// --- Siemens Structured Format ---
DATA_BLOCK "model__HS32_IW100_"
{ S7_Optimized_Access := 'TRUE' }
VERSION :
NON_RETAIN
   VAR
      W_i : ARRAY[0..31, 0..39] OF REAL;
      W_f : ARRAY[0..31, 0..39] OF REAL;
      W_g : ARRAY[0..31, 0..39] OF REAL;
      W_o : ARRAY[0..31, 0..39] OF REAL;
      R_i : ARRAY[0..31, 0..31] OF REAL;
      R_f : ARRAY[0..31, 0..31] OF REAL;
      R_g : ARRAY[0..31, 0..31] OF REAL;
      R_o : ARRAY[0..31, 0..31] OF REAL;
      B_i : ARRAY[0..31] OF REAL;
      B_f : ARRAY[0..31] OF REAL;
      B_g : ARRAY[0..31] OF REAL;
      B_o : ARRAY[0..31] OF REAL;
      FC_W : ARRAY[0..39, 0..31] OF REAL;
      FC_B : ARRAY[0..39] OF REAL;
   END_VAR
BEGIN

      W_i[0,0] := 0.06179943;
      W_i[0,1] := 0.02775717;
      W_i[0,2] := -0.03196508;
      W_i[0,3] := 0.03677268;
      W_i[0,4] := 0.05541879;
      W_i[0,5] := -0.02846526;
      W_i[0,6] := 0.05010877;
      W_i[0,7] := 0.04675795;
      W_i[0,8] := 0.08269168;
      W_i[0,9] := -0.01895206;
      W_i[0,10] := 0.01859271;
      W_i[0,11] := -0.13412605;
      W_i[0,12] := 0.22322017;
      W_i[0,13] := 0.00698021;
      W_i[0,14] := 0.01548957;
      W_i[0,15] := -0.04365166;
      W_i[0,16] := -0.03781708;
      W_i[0,17] := 0.00911400;
      W_i[0,18] := -0.02057064;
      W_i[0,19] := -0.08685457;
      W_i[0,20] := -0.01680454;
      W_i[0,21] := -0.04614456;
      W_i[0,22] := -0.03545121;
      W_i[0,23] := -0.02339789;
      W_i[0,24] := -1.12611961;
      W_i[0,25] := -0.10453429;
      W_i[0,26] := -0.07026759;
      W_i[0,27] := -0.05480277;
      W_i[0,28] := -0.02404995;
      W_i[0,29] := 0.12750483;
      W_i[0,30] := 0.17675591;
      W_i[0,31] := -0.02635767;
      W_i[0,32] := 0.19571228;
      W_i[0,33] := 0.06735895;
      W_i[0,34] := -0.14900623;
      W_i[0,35] := 0.06775700;
      W_i[0,36] := -0.00490537;
      W_i[0,37] := -0.01378909;
      W_i[0,38] := 0.07458769;
      W_i[0,39] := 0.66414231;
      W_i[1,0] := 0.02071806;
      W_i[1,1] := -0.03353070;
      W_i[1,2] := -0.01928122;
      W_i[1,3] := 0.06214599;
      W_i[1,4] := 0.25778303;
      W_i[1,5] := 0.16688786;
      W_i[1,6] := 0.11954694;
      W_i[1,7] := 0.06900051;
      W_i[1,8] := 0.01723209;
      W_i[1,9] := -0.11005860;
      W_i[1,10] := -0.04237102;
      W_i[1,11] := 0.01513118;
      W_i[1,12] := -0.15226158;
      W_i[1,13] := 0.03596478;
      W_i[1,14] := 0.02140439;
      W_i[1,15] := 0.06197662;
      W_i[1,16] := 0.00865395;
      W_i[1,17] := 0.04867539;
      W_i[1,18] := 0.04397345;
      W_i[1,19] := 0.06557351;
      W_i[1,20] := 0.06942460;
      W_i[1,21] := 0.05065425;
      W_i[1,22] := 0.10510546;
      W_i[1,23] := 0.04281416;
      W_i[1,24] := -0.29392853;
      W_i[1,25] := -0.38343686;
      W_i[1,26] := -0.10036848;
      W_i[1,27] := -0.04264174;
      W_i[1,28] := -0.17839937;
      W_i[1,29] := -0.21495967;
      W_i[1,30] := -0.22097401;
      W_i[1,31] := 0.03829467;
      W_i[1,32] := -0.31760472;
      W_i[1,33] := -0.17684405;
      W_i[1,34] := -0.23336750;
      W_i[1,35] := -0.15993148;
      W_i[1,36] := -0.00517801;
      W_i[1,37] := -0.01187338;
      W_i[1,38] := -0.03392988;
      W_i[1,39] := -0.04533037;
      W_i[2,0] := -0.00829509;
      W_i[2,1] := -0.14865589;
      W_i[2,2] := -0.01495113;
      W_i[2,3] := 0.02128208;
      W_i[2,4] := 0.21340890;
      W_i[2,5] := -0.05039188;
      W_i[2,6] := 0.02410355;
      W_i[2,7] := -0.16800745;
      W_i[2,8] := -0.07282868;
      W_i[2,9] := -0.06157869;
      W_i[2,10] := 0.17263004;
      W_i[2,11] := 0.02063438;
      W_i[2,12] := 0.17519112;
      W_i[2,13] := -0.00622400;
      W_i[2,14] := 0.06819141;
      W_i[2,15] := 0.06226488;
      W_i[2,16] := -0.03465794;
      W_i[2,17] := 0.02215759;
      W_i[2,18] := -0.05341673;
      W_i[2,19] := -0.13253070;
      W_i[2,20] := 0.04460967;
      W_i[2,21] := 0.11263417;
      W_i[2,22] := 0.09742771;
      W_i[2,23] := 0.00662358;
      W_i[2,24] := -0.05392387;
      W_i[2,25] := -0.17852309;
      W_i[2,26] := 0.03923597;
      W_i[2,27] := -0.02955864;
      W_i[2,28] := 0.03645090;
      W_i[2,29] := -0.03638797;
      W_i[2,30] := 0.33836386;
      W_i[2,31] := 0.12495890;
      W_i[2,32] := 0.06078594;
      W_i[2,33] := -0.14091927;
      W_i[2,34] := 0.17067178;
      W_i[2,35] := -0.12043836;
      W_i[2,36] := -0.01742014;
      W_i[2,37] := -0.29951882;
      W_i[2,38] := 0.04487922;
      W_i[2,39] := -0.04771054;
      W_i[3,0] := -0.00100313;
      W_i[3,1] := -0.00449658;
      W_i[3,2] := -0.07554256;
      W_i[3,3] := -0.18185882;
      W_i[3,4] := -0.02607848;
      W_i[3,5] := -0.07896423;
      W_i[3,6] := 0.05784221;
      W_i[3,7] := -0.07038090;
      W_i[3,8] := 0.20566469;
      W_i[3,9] := 0.09180041;
      W_i[3,10] := 0.05098312;
      W_i[3,11] := 0.15374708;
      W_i[3,12] := -0.45315537;
      W_i[3,13] := 0.08420219;
      W_i[3,14] := -0.12126628;
      W_i[3,15] := -0.08021345;
      W_i[3,16] := -0.27470666;
      W_i[3,17] := 0.07300078;
      W_i[3,18] := 0.22311375;
      W_i[3,19] := -0.02914955;
      W_i[3,20] := -0.01066327;
      W_i[3,21] := -0.00681991;
      W_i[3,22] := 0.24156007;
      W_i[3,23] := -0.11151634;
      W_i[3,24] := -0.08966236;
      W_i[3,25] := 0.01983345;
      W_i[3,26] := -0.08444024;
      W_i[3,27] := 0.16410163;
      W_i[3,28] := -0.04299213;
      W_i[3,29] := -0.12410518;
      W_i[3,30] := 0.26584405;
      W_i[3,31] := -0.29169789;
      W_i[3,32] := 0.05328545;
      W_i[3,33] := -0.51094949;
      W_i[3,34] := 0.03447641;
      W_i[3,35] := 0.00506896;
      W_i[3,36] := 0.03782123;
      W_i[3,37] := 0.18697615;
      W_i[3,38] := 0.00981322;
      W_i[3,39] := 0.75137496;
      W_i[4,0] := 0.04553370;
      W_i[4,1] := 0.11792795;
      W_i[4,2] := -0.01621435;
      W_i[4,3] := -0.03620827;
      W_i[4,4] := -0.15278673;
      W_i[4,5] := -0.01032144;
      W_i[4,6] := 0.00459723;
      W_i[4,7] := 0.03891215;
      W_i[4,8] := -0.05662930;
      W_i[4,9] := -0.06458510;
      W_i[4,10] := 0.27832294;
      W_i[4,11] := 0.05678938;
      W_i[4,12] := 0.01970386;
      W_i[4,13] := 0.09437083;
      W_i[4,14] := -0.01984982;
      W_i[4,15] := -0.05285306;
      W_i[4,16] := 0.02962786;
      W_i[4,17] := 0.00963242;
      W_i[4,18] := 0.00985712;
      W_i[4,19] := -0.07215877;
      W_i[4,20] := 0.09223086;
      W_i[4,21] := -0.08452385;
      W_i[4,22] := -0.03868546;
      W_i[4,23] := -0.02803059;
      W_i[4,24] := 0.19232845;
      W_i[4,25] := 0.21442333;
      W_i[4,26] := -0.10829803;
      W_i[4,27] := 0.09679998;
      W_i[4,28] := -0.05681482;
      W_i[4,29] := 0.04554670;
      W_i[4,30] := -0.12465099;
      W_i[4,31] := 0.02753920;
      W_i[4,32] := 0.05632669;
      W_i[4,33] := 0.24204549;
      W_i[4,34] := 0.14613600;
      W_i[4,35] := -0.21246302;
      W_i[4,36] := -0.06815854;
      W_i[4,37] := -0.23073821;
      W_i[4,38] := 0.02998499;
      W_i[4,39] := -0.02546969;
      W_i[5,0] := -0.09215746;
      W_i[5,1] := -0.08727002;
      W_i[5,2] := 0.02556904;
      W_i[5,3] := 0.15369390;
      W_i[5,4] := 0.01142898;
      W_i[5,5] := -0.05077455;
      W_i[5,6] := -0.11507938;
      W_i[5,7] := -0.10518788;
      W_i[5,8] := -0.04785325;
      W_i[5,9] := -0.05123279;
      W_i[5,10] := 0.15905567;
      W_i[5,11] := 0.06097380;
      W_i[5,12] := -0.18418492;
      W_i[5,13] := -0.03047887;
      W_i[5,14] := 0.11933848;
      W_i[5,15] := -0.03554063;
      W_i[5,16] := -0.07242216;
      W_i[5,17] := 0.02859983;
      W_i[5,18] := -0.03490715;
      W_i[5,19] := 0.05818025;
      W_i[5,20] := -0.07515050;
      W_i[5,21] := 0.02579406;
      W_i[5,22] := -0.31216845;
      W_i[5,23] := 0.04713825;
      W_i[5,24] := -0.20269118;
      W_i[5,25] := 0.10239060;
      W_i[5,26] := -0.01558112;
      W_i[5,27] := 0.00159392;
      W_i[5,28] := -0.05441242;
      W_i[5,29] := 0.52095068;
      W_i[5,30] := -0.57061511;
      W_i[5,31] := 0.13902861;
      W_i[5,32] := -0.12816451;
      W_i[5,33] := 0.06774098;
      W_i[5,34] := -0.41744006;
      W_i[5,35] := 0.05064213;
      W_i[5,36] := -0.09991191;
      W_i[5,37] := -0.17586561;
      W_i[5,38] := 0.19242531;
      W_i[5,39] := 0.03359242;
      W_i[6,0] := -0.03353223;
      W_i[6,1] := 0.00677240;
      W_i[6,2] := -0.01104784;
      W_i[6,3] := 0.07707670;
      W_i[6,4] := 0.00404718;
      W_i[6,5] := -0.05442240;
      W_i[6,6] := 0.10070097;
      W_i[6,7] := 0.04808670;
      W_i[6,8] := -0.10168398;
      W_i[6,9] := -0.02940839;
      W_i[6,10] := 0.04046509;
      W_i[6,11] := -0.12609679;
      W_i[6,12] := -0.11311707;
      W_i[6,13] := 0.04389359;
      W_i[6,14] := 0.01754723;
      W_i[6,15] := 0.03694800;
      W_i[6,16] := -0.09526791;
      W_i[6,17] := -0.13010779;
      W_i[6,18] := 0.31546634;
      W_i[6,19] := -0.07569441;
      W_i[6,20] := 0.28956288;
      W_i[6,21] := 0.00949547;
      W_i[6,22] := 0.09859776;
      W_i[6,23] := -0.02917805;
      W_i[6,24] := 0.17138363;
      W_i[6,25] := 0.27182287;
      W_i[6,26] := 0.01862298;
      W_i[6,27] := -0.00405888;
      W_i[6,28] := 0.07469607;
      W_i[6,29] := -0.15340948;
      W_i[6,30] := 0.13516009;
      W_i[6,31] := -0.14186700;
      W_i[6,32] := 0.17514557;
      W_i[6,33] := 0.08133219;
      W_i[6,34] := 0.32842028;
      W_i[6,35] := -0.12072788;
      W_i[6,36] := -0.05676087;
      W_i[6,37] := -0.11963397;
      W_i[6,38] := 0.00256419;
      W_i[6,39] := 0.28269264;
      W_i[7,0] := -0.14775136;
      W_i[7,1] := -0.12126163;
      W_i[7,2] := -0.01920290;
      W_i[7,3] := 0.25063628;
      W_i[7,4] := -0.02222757;
      W_i[7,5] := -0.03862220;
      W_i[7,6] := -0.13837403;
      W_i[7,7] := 0.38717154;
      W_i[7,8] := -0.11613367;
      W_i[7,9] := -0.53373992;
      W_i[7,10] := -0.09174719;
      W_i[7,11] := -0.12254320;
      W_i[7,12] := -0.00825407;
      W_i[7,13] := -0.05826338;
      W_i[7,14] := 0.09619932;
      W_i[7,15] := 0.07305111;
      W_i[7,16] := -0.07672185;
      W_i[7,17] := 0.01172826;
      W_i[7,18] := 0.43864861;
      W_i[7,19] := 0.05868300;
      W_i[7,20] := 0.02254522;
      W_i[7,21] := -0.00708780;
      W_i[7,22] := -0.17880507;
      W_i[7,23] := 0.03120665;
      W_i[7,24] := -0.34886146;
      W_i[7,25] := -0.04237240;
      W_i[7,26] := 0.11693397;
      W_i[7,27] := 0.06307583;
      W_i[7,28] := -0.04923550;
      W_i[7,29] := 0.30479616;
      W_i[7,30] := -0.03511298;
      W_i[7,31] := -0.07993785;
      W_i[7,32] := -0.19723724;
      W_i[7,33] := 0.09875282;
      W_i[7,34] := 0.06003888;
      W_i[7,35] := 0.01167319;
      W_i[7,36] := 0.01233812;
      W_i[7,37] := 0.13565342;
      W_i[7,38] := 0.07438924;
      W_i[7,39] := -0.04580714;
      W_i[8,0] := -0.20123592;
      W_i[8,1] := -0.01675500;
      W_i[8,2] := 0.06737890;
      W_i[8,3] := -0.03567418;
      W_i[8,4] := 0.03670733;
      W_i[8,5] := 0.00518049;
      W_i[8,6] := -0.05625178;
      W_i[8,7] := -0.21017089;
      W_i[8,8] := 0.02617608;
      W_i[8,9] := 0.21776345;
      W_i[8,10] := 0.04046187;
      W_i[8,11] := 0.01215424;
      W_i[8,12] := -0.13758895;
      W_i[8,13] := -0.03766741;
      W_i[8,14] := -0.10688125;
      W_i[8,15] := -0.03897357;
      W_i[8,16] := -0.04154058;
      W_i[8,17] := -0.04646260;
      W_i[8,18] := -0.01917167;
      W_i[8,19] := 0.05721129;
      W_i[8,20] := -0.05588107;
      W_i[8,21] := -0.07682938;
      W_i[8,22] := -0.07860053;
      W_i[8,23] := -0.06132534;
      W_i[8,24] := 0.03326328;
      W_i[8,25] := 0.08150295;
      W_i[8,26] := -0.14111993;
      W_i[8,27] := 0.00011063;
      W_i[8,28] := 0.01932795;
      W_i[8,29] := 0.04262755;
      W_i[8,30] := 0.05650154;
      W_i[8,31] := -0.15539150;
      W_i[8,32] := 0.17859717;
      W_i[8,33] := 0.01948488;
      W_i[8,34] := 0.08800947;
      W_i[8,35] := 0.09776416;
      W_i[8,36] := -0.05269374;
      W_i[8,37] := 0.06550130;
      W_i[8,38] := -0.08607090;
      W_i[8,39] := 0.15070331;
      W_i[9,0] := -0.27159375;
      W_i[9,1] := -0.02797615;
      W_i[9,2] := -0.00100640;
      W_i[9,3] := 0.12800276;
      W_i[9,4] := -0.09242823;
      W_i[9,5] := 0.01892278;
      W_i[9,6] := -0.02738959;
      W_i[9,7] := 0.09567204;
      W_i[9,8] := -0.44594380;
      W_i[9,9] := 0.20733841;
      W_i[9,10] := -0.07766859;
      W_i[9,11] := -0.13440070;
      W_i[9,12] := 0.01596364;
      W_i[9,13] := 0.07334067;
      W_i[9,14] := 0.07882207;
      W_i[9,15] := 0.05607220;
      W_i[9,16] := -0.07642873;
      W_i[9,17] := 0.08819333;
      W_i[9,18] := 0.02835996;
      W_i[9,19] := 0.09605386;
      W_i[9,20] := 0.12935719;
      W_i[9,21] := -0.04795177;
      W_i[9,22] := -0.05849212;
      W_i[9,23] := -0.00860680;
      W_i[9,24] := -0.05882631;
      W_i[9,25] := 0.12313552;
      W_i[9,26] := -0.10078515;
      W_i[9,27] := 0.10558646;
      W_i[9,28] := 0.04912272;
      W_i[9,29] := -0.09551237;
      W_i[9,30] := -0.09409142;
      W_i[9,31] := -0.22199608;
      W_i[9,32] := 0.08531553;
      W_i[9,33] := -0.01295959;
      W_i[9,34] := 0.28744900;
      W_i[9,35] := -0.14239824;
      W_i[9,36] := -0.16849788;
      W_i[9,37] := -0.06152735;
      W_i[9,38] := 0.01881091;
      W_i[9,39] := -0.08872003;
      W_i[10,0] := 0.04977950;
      W_i[10,1] := 0.01497823;
      W_i[10,2] := -0.00536506;
      W_i[10,3] := 0.02952771;
      W_i[10,4] := -0.03139960;
      W_i[10,5] := -0.00463935;
      W_i[10,6] := -0.10389712;
      W_i[10,7] := -0.10033682;
      W_i[10,8] := 0.11073951;
      W_i[10,9] := -0.08885644;
      W_i[10,10] := 0.01201617;
      W_i[10,11] := -0.63600385;
      W_i[10,12] := 0.57826489;
      W_i[10,13] := -0.00285191;
      W_i[10,14] := -0.13222906;
      W_i[10,15] := 0.01793578;
      W_i[10,16] := -0.03972865;
      W_i[10,17] := 0.16141385;
      W_i[10,18] := 0.48685026;
      W_i[10,19] := -0.04842542;
      W_i[10,20] := 0.03557721;
      W_i[10,21] := -0.02083956;
      W_i[10,22] := 0.07665567;
      W_i[10,23] := 0.13016869;
      W_i[10,24] := -0.08724608;
      W_i[10,25] := -0.20036544;
      W_i[10,26] := -0.12496603;
      W_i[10,27] := -0.05189490;
      W_i[10,28] := 0.10159702;
      W_i[10,29] := -0.05331298;
      W_i[10,30] := 0.03033962;
      W_i[10,31] := 0.07102174;
      W_i[10,32] := 0.02948349;
      W_i[10,33] := 0.01139331;
      W_i[10,34] := -0.43736589;
      W_i[10,35] := 0.28173751;
      W_i[10,36] := 0.01866223;
      W_i[10,37] := 0.25957814;
      W_i[10,38] := 0.14778605;
      W_i[10,39] := 0.93045533;
      W_i[11,0] := -0.10133153;
      W_i[11,1] := -0.05051550;
      W_i[11,2] := -0.03669089;
      W_i[11,3] := 0.14228435;
      W_i[11,4] := 0.08680110;
      W_i[11,5] := 0.02299375;
      W_i[11,6] := -0.11019665;
      W_i[11,7] := 0.03878751;
      W_i[11,8] := 0.05327412;
      W_i[11,9] := -0.29215959;
      W_i[11,10] := -0.06103910;
      W_i[11,11] := -0.04436091;
      W_i[11,12] := 0.10810567;
      W_i[11,13] := -0.12327234;
      W_i[11,14] := -0.03792057;
      W_i[11,15] := -0.01659554;
      W_i[11,16] := 0.01878507;
      W_i[11,17] := -0.00647482;
      W_i[11,18] := -0.04410561;
      W_i[11,19] := 0.07929806;
      W_i[11,20] := 0.01020784;
      W_i[11,21] := 0.08437648;
      W_i[11,22] := 0.10375391;
      W_i[11,23] := 0.20762387;
      W_i[11,24] := -0.57340568;
      W_i[11,25] := -0.59531760;
      W_i[11,26] := -0.17425776;
      W_i[11,27] := -0.11098373;
      W_i[11,28] := 0.01483229;
      W_i[11,29] := 0.08123992;
      W_i[11,30] := 0.16729805;
      W_i[11,31] := -0.17426890;
      W_i[11,32] := 0.17722335;
      W_i[11,33] := -0.07652548;
      W_i[11,34] := 0.18267493;
      W_i[11,35] := 0.19876397;
      W_i[11,36] := 0.04698262;
      W_i[11,37] := 0.02095936;
      W_i[11,38] := -0.10085329;
      W_i[11,39] := 1.06740248;
      W_i[12,0] := -0.12894745;
      W_i[12,1] := -0.01604900;
      W_i[12,2] := -0.05750192;
      W_i[12,3] := 0.08071270;
      W_i[12,4] := -0.10707285;
      W_i[12,5] := -0.09226165;
      W_i[12,6] := 0.01451022;
      W_i[12,7] := 0.16588750;
      W_i[12,8] := -0.20528767;
      W_i[12,9] := 0.16444704;
      W_i[12,10] := 0.09167138;
      W_i[12,11] := -0.05738107;
      W_i[12,12] := -0.03085519;
      W_i[12,13] := 0.02227092;
      W_i[12,14] := 0.00619229;
      W_i[12,15] := 0.07799102;
      W_i[12,16] := 0.02899228;
      W_i[12,17] := 0.01908563;
      W_i[12,18] := 0.55716008;
      W_i[12,19] := 0.09226023;
      W_i[12,20] := -0.01587960;
      W_i[12,21] := -0.13448635;
      W_i[12,22] := -0.14700012;
      W_i[12,23] := -0.06094320;
      W_i[12,24] := 0.27282214;
      W_i[12,25] := 0.21529709;
      W_i[12,26] := -0.12392846;
      W_i[12,27] := 0.05751082;
      W_i[12,28] := 0.12284551;
      W_i[12,29] := -0.00490399;
      W_i[12,30] := -0.17141145;
      W_i[12,31] := -0.08434223;
      W_i[12,32] := 0.05438624;
      W_i[12,33] := -0.10759345;
      W_i[12,34] := -0.07436828;
      W_i[12,35] := -0.12592168;
      W_i[12,36] := 0.02604092;
      W_i[12,37] := -0.15142396;
      W_i[12,38] := -0.03170886;
      W_i[12,39] := 0.16621175;
      W_i[13,0] := -0.00913993;
      W_i[13,1] := -0.04174744;
      W_i[13,2] := -0.03129856;
      W_i[13,3] := -0.04003599;
      W_i[13,4] := 0.04255468;
      W_i[13,5] := 0.00480728;
      W_i[13,6] := -0.07061405;
      W_i[13,7] := -0.03280373;
      W_i[13,8] := 0.02827574;
      W_i[13,9] := 0.02418965;
      W_i[13,10] := 0.07189363;
      W_i[13,11] := 0.12613529;
      W_i[13,12] := 0.03361855;
      W_i[13,13] := 0.03988501;
      W_i[13,14] := -0.02885863;
      W_i[13,15] := -0.00470651;
      W_i[13,16] := -0.03359226;
      W_i[13,17] := -0.00056631;
      W_i[13,18] := -0.07915758;
      W_i[13,19] := 0.01315921;
      W_i[13,20] := 0.10718971;
      W_i[13,21] := 0.13062805;
      W_i[13,22] := 0.16784896;
      W_i[13,23] := -0.07162543;
      W_i[13,24] := 0.03916876;
      W_i[13,25] := -0.11025614;
      W_i[13,26] := -0.04175865;
      W_i[13,27] := -0.27723673;
      W_i[13,28] := 0.18863167;
      W_i[13,29] := 0.18414941;
      W_i[13,30] := 0.21448347;
      W_i[13,31] := 0.27937597;
      W_i[13,32] := -0.15358151;
      W_i[13,33] := 0.04613268;
      W_i[13,34] := -0.28416333;
      W_i[13,35] := -0.24947314;
      W_i[13,36] := -0.06312902;
      W_i[13,37] := -0.19301520;
      W_i[13,38] := 0.07415584;
      W_i[13,39] := 0.07214847;
      W_i[14,0] := -0.06886686;
      W_i[14,1] := 0.09983595;
      W_i[14,2] := 0.00539746;
      W_i[14,3] := 0.03236075;
      W_i[14,4] := 0.30145952;
      W_i[14,5] := 0.10646193;
      W_i[14,6] := -0.00687617;
      W_i[14,7] := -0.02083724;
      W_i[14,8] := 0.09362940;
      W_i[14,9] := 0.24021219;
      W_i[14,10] := -0.51702040;
      W_i[14,11] := 0.00785133;
      W_i[14,12] := -0.06570137;
      W_i[14,13] := 0.00066462;
      W_i[14,14] := 0.04833549;
      W_i[14,15] := 0.01324825;
      W_i[14,16] := 0.00547472;
      W_i[14,17] := 0.03968929;
      W_i[14,18] := -0.05878792;
      W_i[14,19] := -0.12701105;
      W_i[14,20] := 0.64508420;
      W_i[14,21] := -0.02393116;
      W_i[14,22] := 0.01463204;
      W_i[14,23] := 0.09599538;
      W_i[14,24] := -0.01352467;
      W_i[14,25] := -0.09434310;
      W_i[14,26] := 0.09360847;
      W_i[14,27] := 0.19543391;
      W_i[14,28] := -0.08615168;
      W_i[14,29] := 0.51883084;
      W_i[14,30] := 0.05632273;
      W_i[14,31] := 0.31189725;
      W_i[14,32] := -0.08525938;
      W_i[14,33] := 0.18389013;
      W_i[14,34] := 0.22316632;
      W_i[14,35] := -0.11821964;
      W_i[14,36] := 0.02146083;
      W_i[14,37] := -0.16101155;
      W_i[14,38] := 0.00918483;
      W_i[14,39] := -0.08109198;
      W_i[15,0] := 0.08172593;
      W_i[15,1] := -0.15062873;
      W_i[15,2] := 0.00789237;
      W_i[15,3] := -0.12266801;
      W_i[15,4] := -0.01449642;
      W_i[15,5] := -0.08026960;
      W_i[15,6] := 0.00158959;
      W_i[15,7] := -0.17118339;
      W_i[15,8] := 0.06299323;
      W_i[15,9] := 0.08208384;
      W_i[15,10] := 0.04913726;
      W_i[15,11] := -0.04209859;
      W_i[15,12] := 0.14104722;
      W_i[15,13] := 0.08269731;
      W_i[15,14] := -0.00785436;
      W_i[15,15] := 0.01761792;
      W_i[15,16] := 0.06018753;
      W_i[15,17] := 0.01103730;
      W_i[15,18] := 0.60089856;
      W_i[15,19] := -0.02956709;
      W_i[15,20] := -0.06978408;
      W_i[15,21] := -0.10184263;
      W_i[15,22] := -0.08161820;
      W_i[15,23] := -0.09385420;
      W_i[15,24] := -0.25269318;
      W_i[15,25] := -0.36792046;
      W_i[15,26] := -0.02104633;
      W_i[15,27] := 0.08724175;
      W_i[15,28] := -0.02899375;
      W_i[15,29] := 0.06102180;
      W_i[15,30] := -0.07059706;
      W_i[15,31] := 0.02143796;
      W_i[15,32] := -0.10914523;
      W_i[15,33] := -0.00082962;
      W_i[15,34] := -0.13892201;
      W_i[15,35] := 0.03998528;
      W_i[15,36] := -0.00446972;
      W_i[15,37] := 0.06410963;
      W_i[15,38] := -0.09802709;
      W_i[15,39] := 0.13650982;
      W_i[16,0] := 0.00692594;
      W_i[16,1] := -0.06901163;
      W_i[16,2] := -0.06960113;
      W_i[16,3] := 0.01490095;
      W_i[16,4] := 0.11437556;
      W_i[16,5] := -0.10528261;
      W_i[16,6] := 0.06423379;
      W_i[16,7] := -0.09478712;
      W_i[16,8] := -0.00620357;
      W_i[16,9] := 0.04550839;
      W_i[16,10] := 0.06371807;
      W_i[16,11] := -0.22288436;
      W_i[16,12] := 0.11317084;
      W_i[16,13] := -0.00150014;
      W_i[16,14] := 0.03941125;
      W_i[16,15] := 0.23517418;
      W_i[16,16] := 0.06774591;
      W_i[16,17] := -0.06179966;
      W_i[16,18] := -0.02661809;
      W_i[16,19] := -0.46718821;
      W_i[16,20] := 0.00290592;
      W_i[16,21] := 0.08730330;
      W_i[16,22] := -0.17280819;
      W_i[16,23] := 0.04183443;
      W_i[16,24] := -0.15965074;
      W_i[16,25] := -0.21877262;
      W_i[16,26] := 0.03479860;
      W_i[16,27] := -0.03698987;
      W_i[16,28] := -0.04753701;
      W_i[16,29] := 0.12801097;
      W_i[16,30] := 0.04739811;
      W_i[16,31] := -0.00796509;
      W_i[16,32] := -0.10788697;
      W_i[16,33] := -0.08236082;
      W_i[16,34] := -0.41695821;
      W_i[16,35] := 0.02638846;
      W_i[16,36] := -0.05947839;
      W_i[16,37] := -0.08056837;
      W_i[16,38] := 0.04219051;
      W_i[16,39] := -0.06786148;
      W_i[17,0] := 0.19944434;
      W_i[17,1] := 0.11471956;
      W_i[17,2] := 0.00180160;
      W_i[17,3] := 0.11797725;
      W_i[17,4] := -0.12125240;
      W_i[17,5] := 0.27995679;
      W_i[17,6] := -0.34394604;
      W_i[17,7] := 0.02910547;
      W_i[17,8] := -0.19582599;
      W_i[17,9] := -0.11236304;
      W_i[17,10] := -0.31493005;
      W_i[17,11] := -0.24195738;
      W_i[17,12] := -0.07686605;
      W_i[17,13] := 0.14992486;
      W_i[17,14] := -0.19373207;
      W_i[17,15] := -0.25997469;
      W_i[17,16] := 0.04234881;
      W_i[17,17] := -0.07211331;
      W_i[17,18] := 0.13888460;
      W_i[17,19] := -0.12404422;
      W_i[17,20] := -0.08650170;
      W_i[17,21] := 0.22232069;
      W_i[17,22] := 0.02460083;
      W_i[17,23] := -0.23321719;
      W_i[17,24] := 0.27493891;
      W_i[17,25] := 0.29532185;
      W_i[17,26] := -0.09839682;
      W_i[17,27] := -0.27084854;
      W_i[17,28] := 0.16536197;
      W_i[17,29] := 0.96769738;
      W_i[17,30] := 0.08850956;
      W_i[17,31] := 0.44717026;
      W_i[17,32] := 0.05195052;
      W_i[17,33] := -0.25492772;
      W_i[17,34] := 0.08993755;
      W_i[17,35] := 0.11916504;
      W_i[17,36] := 0.51604098;
      W_i[17,37] := -0.19514880;
      W_i[17,38] := 0.03904369;
      W_i[17,39] := -1.25412786;
      W_i[18,0] := 0.26778793;
      W_i[18,1] := -0.01803258;
      W_i[18,2] := -0.35264796;
      W_i[18,3] := -0.03628552;
      W_i[18,4] := -0.09051698;
      W_i[18,5] := -0.07353226;
      W_i[18,6] := -0.03659349;
      W_i[18,7] := 0.01280040;
      W_i[18,8] := -0.03461934;
      W_i[18,9] := 0.05958343;
      W_i[18,10] := 0.05166731;
      W_i[18,11] := -0.09699293;
      W_i[18,12] := -0.12538935;
      W_i[18,13] := -0.00645365;
      W_i[18,14] := 0.02199500;
      W_i[18,15] := -0.03021014;
      W_i[18,16] := 0.18712366;
      W_i[18,17] := -0.01909142;
      W_i[18,18] := 0.02058483;
      W_i[18,19] := 0.08988243;
      W_i[18,20] := 0.07572187;
      W_i[18,21] := 0.08197203;
      W_i[18,22] := -0.07564746;
      W_i[18,23] := 0.03924798;
      W_i[18,24] := -0.40492132;
      W_i[18,25] := -0.37123427;
      W_i[18,26] := 0.04573231;
      W_i[18,27] := -0.01739427;
      W_i[18,28] := -0.00431714;
      W_i[18,29] := 0.16991295;
      W_i[18,30] := -0.03938163;
      W_i[18,31] := -0.01546910;
      W_i[18,32] := -0.25745204;
      W_i[18,33] := 0.13622859;
      W_i[18,34] := -0.16286966;
      W_i[18,35] := -0.25323087;
      W_i[18,36] := 0.02914849;
      W_i[18,37] := 0.00573681;
      W_i[18,38] := -0.05729824;
      W_i[18,39] := 0.23888165;
      W_i[19,0] := -0.05738360;
      W_i[19,1] := 0.05517812;
      W_i[19,2] := -0.01163843;
      W_i[19,3] := -0.07037261;
      W_i[19,4] := -0.07145417;
      W_i[19,5] := 0.08916121;
      W_i[19,6] := -0.05329772;
      W_i[19,7] := -0.17612284;
      W_i[19,8] := -0.03184425;
      W_i[19,9] := 0.03378281;
      W_i[19,10] := 0.06813814;
      W_i[19,11] := 0.08680203;
      W_i[19,12] := -0.17591415;
      W_i[19,13] := -0.04395442;
      W_i[19,14] := 0.10378881;
      W_i[19,15] := 0.11948365;
      W_i[19,16] := -0.11327706;
      W_i[19,17] := 0.03809229;
      W_i[19,18] := 0.04363121;
      W_i[19,19] := -0.08202547;
      W_i[19,20] := 0.04668652;
      W_i[19,21] := -0.06396332;
      W_i[19,22] := -0.11801164;
      W_i[19,23] := 0.00545785;
      W_i[19,24] := 0.19188444;
      W_i[19,25] := 0.15162137;
      W_i[19,26] := -0.08233768;
      W_i[19,27] := 0.10989103;
      W_i[19,28] := 0.06658027;
      W_i[19,29] := -0.12314930;
      W_i[19,30] := -0.29401505;
      W_i[19,31] := -0.02752479;
      W_i[19,32] := -0.06132220;
      W_i[19,33] := -0.22982699;
      W_i[19,34] := -0.23728208;
      W_i[19,35] := -0.25140384;
      W_i[19,36] := -0.05633686;
      W_i[19,37] := -0.18172039;
      W_i[19,38] := 0.11977114;
      W_i[19,39] := -0.16488980;
      W_i[20,0] := -0.01835487;
      W_i[20,1] := -0.04570545;
      W_i[20,2] := 0.04467667;
      W_i[20,3] := -0.07336899;
      W_i[20,4] := 0.02571872;
      W_i[20,5] := -0.01889678;
      W_i[20,6] := -0.02779749;
      W_i[20,7] := 0.08607043;
      W_i[20,8] := 0.01099925;
      W_i[20,9] := -0.00992060;
      W_i[20,10] := -0.01524233;
      W_i[20,11] := 0.21199150;
      W_i[20,12] := 0.01592732;
      W_i[20,13] := -0.01826751;
      W_i[20,14] := -0.10014486;
      W_i[20,15] := 0.00661277;
      W_i[20,16] := 0.01667893;
      W_i[20,17] := 0.02136482;
      W_i[20,18] := 0.03966679;
      W_i[20,19] := -0.07920662;
      W_i[20,20] := 0.06787179;
      W_i[20,21] := 0.42317262;
      W_i[20,22] := -0.33591220;
      W_i[20,23] := -0.00585524;
      W_i[20,24] := 0.09470745;
      W_i[20,25] := 0.15506293;
      W_i[20,26] := -0.30801183;
      W_i[20,27] := -0.33458385;
      W_i[20,28] := -0.08752628;
      W_i[20,29] := 0.35584134;
      W_i[20,30] := -0.20388263;
      W_i[20,31] := -0.01898901;
      W_i[20,32] := -0.41883579;
      W_i[20,33] := -0.54509979;
      W_i[20,34] := -0.31911835;
      W_i[20,35] := 0.02712717;
      W_i[20,36] := -0.01844929;
      W_i[20,37] := 0.01240083;
      W_i[20,38] := -0.24291822;
      W_i[20,39] := -0.17812274;
      W_i[21,0] := 0.12280829;
      W_i[21,1] := -0.07471990;
      W_i[21,2] := -0.05163937;
      W_i[21,3] := -0.22502938;
      W_i[21,4] := 0.00184776;
      W_i[21,5] := -0.01510628;
      W_i[21,6] := 0.13238980;
      W_i[21,7] := -0.09605303;
      W_i[21,8] := 0.05345604;
      W_i[21,9] := 0.25691971;
      W_i[21,10] := 0.00038861;
      W_i[21,11] := -0.01645699;
      W_i[21,12] := -0.07529693;
      W_i[21,13] := -0.01089604;
      W_i[21,14] := 0.07050634;
      W_i[21,15] := -0.01411841;
      W_i[21,16] := -0.09095489;
      W_i[21,17] := -0.02065623;
      W_i[21,18] := 0.05196851;
      W_i[21,19] := 0.80753618;
      W_i[21,20] := -0.02273143;
      W_i[21,21] := 0.03218904;
      W_i[21,22] := 0.16152497;
      W_i[21,23] := -0.01746419;
      W_i[21,24] := 0.70909500;
      W_i[21,25] := 0.95648199;
      W_i[21,26] := 0.13566963;
      W_i[21,27] := 0.11187585;
      W_i[21,28] := 0.08011223;
      W_i[21,29] := -0.13311587;
      W_i[21,30] := 0.02521890;
      W_i[21,31] := 0.09288229;
      W_i[21,32] := 0.16024679;
      W_i[21,33] := 0.04743494;
      W_i[21,34] := -0.09396220;
      W_i[21,35] := 0.12562209;
      W_i[21,36] := 0.04016363;
      W_i[21,37] := 0.29017061;
      W_i[21,38] := 0.02795759;
      W_i[21,39] := 0.36647096;
      W_i[22,0] := 0.06585112;
      W_i[22,1] := -0.07038485;
      W_i[22,2] := 0.03823679;
      W_i[22,3] := 0.13506269;
      W_i[22,4] := 0.06941289;
      W_i[22,5] := -0.08188840;
      W_i[22,6] := -0.00802410;
      W_i[22,7] := 0.00843967;
      W_i[22,8] := 0.03293480;
      W_i[22,9] := 0.00418619;
      W_i[22,10] := -0.18440005;
      W_i[22,11] := -0.07325464;
      W_i[22,12] := -0.14550987;
      W_i[22,13] := -0.08753653;
      W_i[22,14] := 0.04707590;
      W_i[22,15] := 0.02154654;
      W_i[22,16] := -0.05312854;
      W_i[22,17] := -0.00624513;
      W_i[22,18] := -0.05160676;
      W_i[22,19] := 0.08727906;
      W_i[22,20] := 0.02189743;
      W_i[22,21] := 0.08372616;
      W_i[22,22] := 0.26144525;
      W_i[22,23] := 0.16893846;
      W_i[22,24] := -0.15793604;
      W_i[22,25] := -0.13311699;
      W_i[22,26] := -0.11365860;
      W_i[22,27] := 0.00836681;
      W_i[22,28] := -0.09337366;
      W_i[22,29] := -0.01833472;
      W_i[22,30] := -0.04223403;
      W_i[22,31] := -0.05326389;
      W_i[22,32] := 0.19289488;
      W_i[22,33] := 0.05630151;
      W_i[22,34] := 0.27636716;
      W_i[22,35] := -0.09883546;
      W_i[22,36] := 0.07930394;
      W_i[22,37] := -0.02333659;
      W_i[22,38] := 0.02749063;
      W_i[22,39] := -0.01253646;
      W_i[23,0] := 0.01285714;
      W_i[23,1] := -0.01090977;
      W_i[23,2] := -0.12196957;
      W_i[23,3] := 0.08748322;
      W_i[23,4] := -0.04398613;
      W_i[23,5] := -0.13556443;
      W_i[23,6] := 0.02350867;
      W_i[23,7] := -0.11876588;
      W_i[23,8] := 0.10013366;
      W_i[23,9] := 0.02939740;
      W_i[23,10] := -0.09517333;
      W_i[23,11] := 0.11568693;
      W_i[23,12] := -0.36971363;
      W_i[23,13] := -0.06232831;
      W_i[23,14] := 0.02247390;
      W_i[23,15] := 0.01112311;
      W_i[23,16] := -0.05705897;
      W_i[23,17] := 0.06032606;
      W_i[23,18] := 0.32368115;
      W_i[23,19] := -0.10644881;
      W_i[23,20] := -0.04895338;
      W_i[23,21] := 0.09499650;
      W_i[23,22] := -0.10231195;
      W_i[23,23] := -0.01488803;
      W_i[23,24] := -0.22148487;
      W_i[23,25] := -0.02040800;
      W_i[23,26] := 0.18095909;
      W_i[23,27] := -0.01085224;
      W_i[23,28] := 0.08920502;
      W_i[23,29] := 0.30755806;
      W_i[23,30] := -0.21824111;
      W_i[23,31] := -0.06937134;
      W_i[23,32] := 0.14039119;
      W_i[23,33] := 0.22622369;
      W_i[23,34] := -0.10339716;
      W_i[23,35] := 0.05056783;
      W_i[23,36] := -0.01605630;
      W_i[23,37] := 0.21682332;
      W_i[23,38] := 0.91564023;
      W_i[23,39] := 0.60147935;
      W_i[24,0] := -0.06349316;
      W_i[24,1] := -0.06430539;
      W_i[24,2] := 0.04938103;
      W_i[24,3] := 0.02899365;
      W_i[24,4] := 0.02045459;
      W_i[24,5] := -0.03727232;
      W_i[24,6] := 0.01954682;
      W_i[24,7] := -0.10346385;
      W_i[24,8] := 0.00335618;
      W_i[24,9] := -0.11790799;
      W_i[24,10] := 0.04728369;
      W_i[24,11] := 0.09648414;
      W_i[24,12] := -0.04300074;
      W_i[24,13] := 0.02185826;
      W_i[24,14] := 0.01268934;
      W_i[24,15] := -0.03640975;
      W_i[24,16] := -0.00692598;
      W_i[24,17] := -0.01243239;
      W_i[24,18] := 0.02085917;
      W_i[24,19] := 0.02911621;
      W_i[24,20] := 0.11124941;
      W_i[24,21] := 0.14329974;
      W_i[24,22] := 0.07946618;
      W_i[24,23] := 0.01397222;
      W_i[24,24] := -0.33342758;
      W_i[24,25] := -0.18193676;
      W_i[24,26] := -0.12712136;
      W_i[24,27] := -0.03829253;
      W_i[24,28] := 0.01048399;
      W_i[24,29] := -0.12682118;
      W_i[24,30] := 0.06314925;
      W_i[24,31] := 0.08736062;
      W_i[24,32] := -0.07333044;
      W_i[24,33] := -0.18093891;
      W_i[24,34] := 0.08127785;
      W_i[24,35] := -0.14450674;
      W_i[24,36] := -0.05644464;
      W_i[24,37] := -0.06005542;
      W_i[24,38] := 0.01570564;
      W_i[24,39] := 0.04107951;
      W_i[25,0] := -0.00392134;
      W_i[25,1] := -0.02218844;
      W_i[25,2] := 0.01908197;
      W_i[25,3] := 0.00515596;
      W_i[25,4] := -0.06599259;
      W_i[25,5] := -0.09139763;
      W_i[25,6] := 0.06393541;
      W_i[25,7] := -0.03314249;
      W_i[25,8] := -0.00094995;
      W_i[25,9] := -0.09238666;
      W_i[25,10] := 0.12895916;
      W_i[25,11] := -0.03478534;
      W_i[25,12] := 0.08731889;
      W_i[25,13] := 0.00909062;
      W_i[25,14] := 0.03396220;
      W_i[25,15] := 0.00441095;
      W_i[25,16] := -0.08805312;
      W_i[25,17] := 0.06228795;
      W_i[25,18] := -0.04030024;
      W_i[25,19] := -0.05294413;
      W_i[25,20] := -0.03475821;
      W_i[25,21] := -0.09267792;
      W_i[25,22] := -0.11669731;
      W_i[25,23] := -0.03766777;
      W_i[25,24] := -0.03449144;
      W_i[25,25] := -0.15750119;
      W_i[25,26] := 0.02700294;
      W_i[25,27] := 0.10468993;
      W_i[25,28] := 0.03980485;
      W_i[25,29] := 0.01171093;
      W_i[25,30] := 0.08682661;
      W_i[25,31] := -0.00671425;
      W_i[25,32] := 0.00725360;
      W_i[25,33] := -0.11579906;
      W_i[25,34] := -0.55428278;
      W_i[25,35] := 0.18704750;
      W_i[25,36] := -0.03766178;
      W_i[25,37] := -0.09676717;
      W_i[25,38] := 0.10681428;
      W_i[25,39] := -0.04854197;
      W_i[26,0] := 0.03223363;
      W_i[26,1] := -0.11389477;
      W_i[26,2] := 0.01710660;
      W_i[26,3] := -0.06687164;
      W_i[26,4] := 0.01613229;
      W_i[26,5] := -0.03883494;
      W_i[26,6] := -0.10788758;
      W_i[26,7] := 0.04997331;
      W_i[26,8] := 0.00840330;
      W_i[26,9] := -0.06306913;
      W_i[26,10] := 0.06178190;
      W_i[26,11] := -0.12198523;
      W_i[26,12] := -0.04752781;
      W_i[26,13] := -0.03431008;
      W_i[26,14] := 0.00714531;
      W_i[26,15] := 0.05213116;
      W_i[26,16] := 0.01167048;
      W_i[26,17] := -0.00677893;
      W_i[26,18] := -0.24137808;
      W_i[26,19] := -0.07195701;
      W_i[26,20] := -0.10280736;
      W_i[26,21] := -0.00431173;
      W_i[26,22] := -0.40525341;
      W_i[26,23] := 0.00794029;
      W_i[26,24] := -0.36122626;
      W_i[26,25] := 0.04784513;
      W_i[26,26] := -0.29187959;
      W_i[26,27] := -0.14297174;
      W_i[26,28] := 0.02196433;
      W_i[26,29] := 0.49258694;
      W_i[26,30] := -0.35673437;
      W_i[26,31] := -0.14768223;
      W_i[26,32] := -0.14340006;
      W_i[26,33] := -0.10875791;
      W_i[26,34] := -0.22464323;
      W_i[26,35] := -0.14221328;
      W_i[26,36] := -0.07692026;
      W_i[26,37] := -0.33565632;
      W_i[26,38] := -0.03680801;
      W_i[26,39] := -0.08500476;
      W_i[27,0] := -0.03908358;
      W_i[27,1] := 0.06247386;
      W_i[27,2] := 0.07315844;
      W_i[27,3] := -0.12355068;
      W_i[27,4] := 0.05118919;
      W_i[27,5] := -0.01427916;
      W_i[27,6] := 0.12830800;
      W_i[27,7] := 0.12413668;
      W_i[27,8] := -0.04524078;
      W_i[27,9] := 0.12099374;
      W_i[27,10] := 0.00551115;
      W_i[27,11] := 0.29388657;
      W_i[27,12] := -0.18307312;
      W_i[27,13] := 0.04645123;
      W_i[27,14] := 0.01536438;
      W_i[27,15] := -0.15575469;
      W_i[27,16] := -0.06600323;
      W_i[27,17] := 0.00907420;
      W_i[27,18] := 0.76988453;
      W_i[27,19] := 0.03355170;
      W_i[27,20] := -0.00380640;
      W_i[27,21] := 0.02491378;
      W_i[27,22] := 0.00787842;
      W_i[27,23] := -0.03097626;
      W_i[27,24] := 0.01564326;
      W_i[27,25] := 0.19453372;
      W_i[27,26] := 0.06244323;
      W_i[27,27] := 0.05636120;
      W_i[27,28] := -0.16548483;
      W_i[27,29] := -0.05327202;
      W_i[27,30] := 0.07400166;
      W_i[27,31] := -0.14070928;
      W_i[27,32] := -0.00810295;
      W_i[27,33] := 0.09415199;
      W_i[27,34] := -0.15936106;
      W_i[27,35] := 0.11152661;
      W_i[27,36] := 0.03231200;
      W_i[27,37] := 0.04753703;
      W_i[27,38] := 0.23126490;
      W_i[27,39] := 0.00431150;
      W_i[28,0] := 0.03881709;
      W_i[28,1] := -0.04091561;
      W_i[28,2] := 0.01611770;
      W_i[28,3] := 0.00697450;
      W_i[28,4] := 0.18305339;
      W_i[28,5] := -0.15279785;
      W_i[28,6] := 0.04542335;
      W_i[28,7] := 0.19088306;
      W_i[28,8] := -0.09130806;
      W_i[28,9] := -0.06414899;
      W_i[28,10] := -0.17731205;
      W_i[28,11] := 0.30202127;
      W_i[28,12] := -0.05439992;
      W_i[28,13] := -0.01150446;
      W_i[28,14] := 0.00131535;
      W_i[28,15] := -0.09205615;
      W_i[28,16] := 0.00188813;
      W_i[28,17] := 0.02027261;
      W_i[28,18] := -0.10595226;
      W_i[28,19] := 0.04467888;
      W_i[28,20] := 0.06951932;
      W_i[28,21] := -0.00705112;
      W_i[28,22] := 0.26304314;
      W_i[28,23] := -0.06421968;
      W_i[28,24] := -0.06970753;
      W_i[28,25] := -0.04688016;
      W_i[28,26] := -0.12970042;
      W_i[28,27] := -0.15225610;
      W_i[28,28] := -0.09705786;
      W_i[28,29] := 0.48931244;
      W_i[28,30] := 0.07042009;
      W_i[28,31] := 0.21406028;
      W_i[28,32] := 0.07373387;
      W_i[28,33] := 0.03300231;
      W_i[28,34] := 0.03395164;
      W_i[28,35] := 0.00114277;
      W_i[28,36] := 0.11038067;
      W_i[28,37] := 0.08363102;
      W_i[28,38] := 0.06231136;
      W_i[28,39] := 0.02984152;
      W_i[29,0] := 0.34138203;
      W_i[29,1] := 0.16524114;
      W_i[29,2] := -0.15652245;
      W_i[29,3] := 0.16650911;
      W_i[29,4] := 0.18447480;
      W_i[29,5] := 0.09144969;
      W_i[29,6] := 0.01847808;
      W_i[29,7] := -0.09755348;
      W_i[29,8] := 0.06849403;
      W_i[29,9] := -0.12883465;
      W_i[29,10] := -0.08249056;
      W_i[29,11] := -0.14052261;
      W_i[29,12] := 0.00471857;
      W_i[29,13] := 0.11108005;
      W_i[29,14] := 0.00168034;
      W_i[29,15] := 0.01264171;
      W_i[29,16] := 0.03052950;
      W_i[29,17] := -0.01635699;
      W_i[29,18] := 0.68267095;
      W_i[29,19] := 0.05182270;
      W_i[29,20] := 0.04084420;
      W_i[29,21] := -0.13725121;
      W_i[29,22] := -0.06725579;
      W_i[29,23] := 0.06445967;
      W_i[29,24] := -0.25235596;
      W_i[29,25] := -0.34174517;
      W_i[29,26] := -0.12284433;
      W_i[29,27] := 0.01959689;
      W_i[29,28] := -0.15510176;
      W_i[29,29] := -0.05445927;
      W_i[29,30] := -0.00391692;
      W_i[29,31] := 0.09164531;
      W_i[29,32] := -0.03895570;
      W_i[29,33] := 0.01729037;
      W_i[29,34] := -0.47271654;
      W_i[29,35] := -0.19013441;
      W_i[29,36] := 0.02730786;
      W_i[29,37] := -0.10548180;
      W_i[29,38] := -0.02444625;
      W_i[29,39] := 0.22114794;
      W_i[30,0] := 0.14259459;
      W_i[30,1] := 0.13030399;
      W_i[30,2] := 0.01574181;
      W_i[30,3] := 0.32909501;
      W_i[30,4] := 0.18247588;
      W_i[30,5] := 0.10201692;
      W_i[30,6] := -0.16793460;
      W_i[30,7] := -0.01608832;
      W_i[30,8] := -0.07945836;
      W_i[30,9] := -0.06400074;
      W_i[30,10] := -0.02339716;
      W_i[30,11] := -0.61556047;
      W_i[30,12] := -0.43913898;
      W_i[30,13] := 0.23748495;
      W_i[30,14] := -0.04515821;
      W_i[30,15] := -0.21111111;
      W_i[30,16] := -0.35755801;
      W_i[30,17] := -0.60449827;
      W_i[30,18] := -0.20390034;
      W_i[30,19] := -0.22386833;
      W_i[30,20] := -0.23623383;
      W_i[30,21] := -0.01274856;
      W_i[30,22] := 0.05771254;
      W_i[30,23] := 0.27973813;
      W_i[30,24] := 0.21776874;
      W_i[30,25] := 0.00964033;
      W_i[30,26] := -0.01853784;
      W_i[30,27] := 0.48116028;
      W_i[30,28] := 0.02131466;
      W_i[30,29] := -0.26301557;
      W_i[30,30] := 0.08809707;
      W_i[30,31] := 0.00659453;
      W_i[30,32] := -0.02935489;
      W_i[30,33] := -0.04626760;
      W_i[30,34] := 0.18829554;
      W_i[30,35] := -0.13441698;
      W_i[30,36] := 0.02834320;
      W_i[30,37] := -0.00632966;
      W_i[30,38] := -0.29868194;
      W_i[30,39] := 0.61415642;
      W_i[31,0] := -0.16325244;
      W_i[31,1] := -0.09679049;
      W_i[31,2] := -0.03050595;
      W_i[31,3] := 0.16190793;
      W_i[31,4] := -0.00247456;
      W_i[31,5] := -0.11562813;
      W_i[31,6] := -0.01968347;
      W_i[31,7] := 0.20883080;
      W_i[31,8] := -0.17580964;
      W_i[31,9] := -0.12375850;
      W_i[31,10] := -0.07372309;
      W_i[31,11] := 0.02056623;
      W_i[31,12] := -0.01187920;
      W_i[31,13] := 0.05266812;
      W_i[31,14] := -0.06564806;
      W_i[31,15] := 0.00189058;
      W_i[31,16] := -0.07726562;
      W_i[31,17] := 0.02975348;
      W_i[31,18] := -0.06461618;
      W_i[31,19] := -0.03122944;
      W_i[31,20] := 0.12285355;
      W_i[31,21] := 0.00985503;
      W_i[31,22] := -0.14180370;
      W_i[31,23] := 0.05783030;
      W_i[31,24] := 0.40578064;
      W_i[31,25] := 0.25383785;
      W_i[31,26] := 0.07038008;
      W_i[31,27] := 0.20337011;
      W_i[31,28] := 0.00104713;
      W_i[31,29] := 0.11606871;
      W_i[31,30] := -0.06506641;
      W_i[31,31] := -0.05263698;
      W_i[31,32] := -0.15003459;
      W_i[31,33] := -0.00927202;
      W_i[31,34] := -0.13444443;
      W_i[31,35] := 0.00383041;
      W_i[31,36] := 0.01434117;
      W_i[31,37] := -0.06329263;
      W_i[31,38] := 0.09013104;
      W_i[31,39] := -0.04022735;
      W_f[0,0] := 0.09275501;
      W_f[0,1] := -0.00732977;
      W_f[0,2] := -0.06869236;
      W_f[0,3] := -0.06190562;
      W_f[0,4] := -0.01295592;
      W_f[0,5] := -0.04590857;
      W_f[0,6] := -0.00253042;
      W_f[0,7] := -0.02688417;
      W_f[0,8] := 0.01320969;
      W_f[0,9] := -0.01583199;
      W_f[0,10] := -0.00835014;
      W_f[0,11] := -0.05974917;
      W_f[0,12] := 0.00843614;
      W_f[0,13] := -0.08353058;
      W_f[0,14] := 0.02314937;
      W_f[0,15] := -0.00417441;
      W_f[0,16] := -0.00421321;
      W_f[0,17] := 0.02465227;
      W_f[0,18] := 0.01412213;
      W_f[0,19] := 0.07288992;
      W_f[0,20] := -0.23401335;
      W_f[0,21] := 0.01645997;
      W_f[0,22] := -0.05039980;
      W_f[0,23] := 0.03279801;
      W_f[0,24] := -0.29735646;
      W_f[0,25] := -0.05838059;
      W_f[0,26] := -0.08404252;
      W_f[0,27] := -0.06417349;
      W_f[0,28] := -0.06763788;
      W_f[0,29] := -0.54978985;
      W_f[0,30] := 0.01095366;
      W_f[0,31] := 0.06258379;
      W_f[0,32] := 0.08439261;
      W_f[0,33] := -0.00216618;
      W_f[0,34] := 0.26842579;
      W_f[0,35] := -0.11115351;
      W_f[0,36] := 0.06083455;
      W_f[0,37] := -0.08760575;
      W_f[0,38] := -0.01485838;
      W_f[0,39] := 0.06713727;
      W_f[1,0] := -0.25717846;
      W_f[1,1] := -0.00925572;
      W_f[1,2] := 0.05973412;
      W_f[1,3] := -0.02157113;
      W_f[1,4] := -0.37918866;
      W_f[1,5] := 0.05476968;
      W_f[1,6] := -0.00041559;
      W_f[1,7] := -0.04717121;
      W_f[1,8] := 0.06120597;
      W_f[1,9] := 0.06802628;
      W_f[1,10] := -0.11830372;
      W_f[1,11] := -0.28673279;
      W_f[1,12] := -0.13959989;
      W_f[1,13] := 0.04275421;
      W_f[1,14] := -0.04769576;
      W_f[1,15] := -0.04396937;
      W_f[1,16] := 0.02418298;
      W_f[1,17] := -0.00998302;
      W_f[1,18] := 0.09016442;
      W_f[1,19] := -0.05595219;
      W_f[1,20] := 0.06755187;
      W_f[1,21] := -0.16743061;
      W_f[1,22] := -0.00463282;
      W_f[1,23] := 0.04815869;
      W_f[1,24] := -0.00236317;
      W_f[1,25] := -0.07198022;
      W_f[1,26] := -0.21302037;
      W_f[1,27] := 0.16784427;
      W_f[1,28] := 0.17687364;
      W_f[1,29] := -0.09877391;
      W_f[1,30] := -0.04312310;
      W_f[1,31] := -0.04830271;
      W_f[1,32] := 0.02740210;
      W_f[1,33] := -0.04927362;
      W_f[1,34] := 0.04876388;
      W_f[1,35] := -0.04135494;
      W_f[1,36] := 0.02199238;
      W_f[1,37] := 0.09235270;
      W_f[1,38] := 0.03114256;
      W_f[1,39] := -0.00403757;
      W_f[2,0] := 0.19074439;
      W_f[2,1] := 0.12946449;
      W_f[2,2] := -0.22353986;
      W_f[2,3] := -0.01812110;
      W_f[2,4] := -0.18054955;
      W_f[2,5] := 0.12059813;
      W_f[2,6] := 0.01315679;
      W_f[2,7] := 0.13689463;
      W_f[2,8] := -0.04521443;
      W_f[2,9] := 0.07877994;
      W_f[2,10] := -0.09594797;
      W_f[2,11] := -0.08541686;
      W_f[2,12] := -0.09018625;
      W_f[2,13] := -0.02363209;
      W_f[2,14] := 0.00390827;
      W_f[2,15] := 0.00712217;
      W_f[2,16] := -0.00533320;
      W_f[2,17] := -0.03277547;
      W_f[2,18] := 0.02854676;
      W_f[2,19] := -0.21850465;
      W_f[2,20] := 0.04750577;
      W_f[2,21] := -0.17764615;
      W_f[2,22] := 0.24915168;
      W_f[2,23] := -0.02141095;
      W_f[2,24] := 1.16149223;
      W_f[2,25] := 0.99568248;
      W_f[2,26] := -0.03115178;
      W_f[2,27] := 0.07513309;
      W_f[2,28] := 0.13894814;
      W_f[2,29] := 0.20039569;
      W_f[2,30] := 0.07511951;
      W_f[2,31] := -0.00536174;
      W_f[2,32] := 0.07269926;
      W_f[2,33] := -0.06267523;
      W_f[2,34] := 1.02267516;
      W_f[2,35] := 0.05643394;
      W_f[2,36] := 0.13621765;
      W_f[2,37] := 0.15765581;
      W_f[2,38] := -0.04730120;
      W_f[2,39] := 0.00392890;
      W_f[3,0] := -0.21518645;
      W_f[3,1] := -0.05239934;
      W_f[3,2] := -0.08921831;
      W_f[3,3] := -0.04948764;
      W_f[3,4] := 0.14105852;
      W_f[3,5] := -0.11283698;
      W_f[3,6] := 0.08679157;
      W_f[3,7] := 0.08755182;
      W_f[3,8] := -0.17906485;
      W_f[3,9] := 0.14633922;
      W_f[3,10] := 0.16945954;
      W_f[3,11] := 0.16170655;
      W_f[3,12] := -0.25333130;
      W_f[3,13] := -0.07672831;
      W_f[3,14] := -0.26473001;
      W_f[3,15] := 0.13318448;
      W_f[3,16] := 0.09231668;
      W_f[3,17] := 0.15904103;
      W_f[3,18] := -0.02022397;
      W_f[3,19] := -0.04273768;
      W_f[3,20] := 0.01525528;
      W_f[3,21] := 0.28678519;
      W_f[3,22] := -0.13602529;
      W_f[3,23] := 0.17240688;
      W_f[3,24] := -0.74654180;
      W_f[3,25] := -0.94593614;
      W_f[3,26] := -0.01936307;
      W_f[3,27] := -0.21515515;
      W_f[3,28] := -0.08529308;
      W_f[3,29] := 0.20380117;
      W_f[3,30] := 0.11490183;
      W_f[3,31] := -0.62479013;
      W_f[3,32] := -0.25840655;
      W_f[3,33] := -0.11416061;
      W_f[3,34] := -1.12916088;
      W_f[3,35] := -0.32786167;
      W_f[3,36] := 0.04079599;
      W_f[3,37] := -0.33860385;
      W_f[3,38] := -0.35431030;
      W_f[3,39] := 1.09083843;
      W_f[4,0] := -0.18852453;
      W_f[4,1] := 0.37211481;
      W_f[4,2] := 0.32904080;
      W_f[4,3] := -0.11470369;
      W_f[4,4] := -0.31123433;
      W_f[4,5] := -0.17510767;
      W_f[4,6] := -0.12685519;
      W_f[4,7] := -0.02077636;
      W_f[4,8] := -0.31811282;
      W_f[4,9] := 0.15811297;
      W_f[4,10] := 0.41503298;
      W_f[4,11] := -0.10261679;
      W_f[4,12] := -0.13673842;
      W_f[4,13] := -0.08312797;
      W_f[4,14] := 0.04571920;
      W_f[4,15] := 0.06901194;
      W_f[4,16] := 0.01600495;
      W_f[4,17] := 0.03952283;
      W_f[4,18] := -0.02872921;
      W_f[4,19] := 0.09338096;
      W_f[4,20] := -0.03377770;
      W_f[4,21] := 0.26424292;
      W_f[4,22] := 0.11843497;
      W_f[4,23] := 0.13067293;
      W_f[4,24] := -0.85125470;
      W_f[4,25] := -0.36451712;
      W_f[4,26] := 0.01728472;
      W_f[4,27] := 0.01718649;
      W_f[4,28] := 0.11088099;
      W_f[4,29] := 0.27615273;
      W_f[4,30] := 0.11448240;
      W_f[4,31] := 0.13193305;
      W_f[4,32] := 0.00523527;
      W_f[4,33] := 0.17511281;
      W_f[4,34] := -0.07963558;
      W_f[4,35] := 0.04655371;
      W_f[4,36] := -0.05894723;
      W_f[4,37] := 0.04638829;
      W_f[4,38] := 0.06854037;
      W_f[4,39] := -0.17245297;
      W_f[5,0] := -0.05104964;
      W_f[5,1] := -0.06627955;
      W_f[5,2] := -0.05809701;
      W_f[5,3] := 0.00228492;
      W_f[5,4] := -0.00232467;
      W_f[5,5] := 0.07671241;
      W_f[5,6] := 0.00179391;
      W_f[5,7] := 0.07644720;
      W_f[5,8] := 0.00137723;
      W_f[5,9] := -0.01465034;
      W_f[5,10] := -0.22236739;
      W_f[5,11] := -0.11612928;
      W_f[5,12] := -0.05232463;
      W_f[5,13] := 0.10474943;
      W_f[5,14] := -0.10528857;
      W_f[5,15] := -0.22751111;
      W_f[5,16] := -0.01253656;
      W_f[5,17] := -0.10420241;
      W_f[5,18] := 0.02031541;
      W_f[5,19] := -0.00450479;
      W_f[5,20] := -0.04310225;
      W_f[5,21] := -0.00651219;
      W_f[5,22] := 0.09841527;
      W_f[5,23] := -0.07680399;
      W_f[5,24] := 0.95654547;
      W_f[5,25] := 0.81427342;
      W_f[5,26] := -0.12573048;
      W_f[5,27] := 0.05082744;
      W_f[5,28] := -0.00532472;
      W_f[5,29] := 0.12227312;
      W_f[5,30] := -0.03822643;
      W_f[5,31] := -0.03150657;
      W_f[5,32] := 0.11010607;
      W_f[5,33] := 0.03363729;
      W_f[5,34] := -0.05923928;
      W_f[5,35] := 0.29333764;
      W_f[5,36] := 0.07078772;
      W_f[5,37] := 0.29227102;
      W_f[5,38] := -0.02658367;
      W_f[5,39] := 0.02677094;
      W_f[6,0] := 0.13546056;
      W_f[6,1] := -0.04973600;
      W_f[6,2] := -0.04891440;
      W_f[6,3] := -0.03705164;
      W_f[6,4] := -0.04525963;
      W_f[6,5] := -0.04312599;
      W_f[6,6] := 0.02302015;
      W_f[6,7] := 0.08248876;
      W_f[6,8] := -0.09446131;
      W_f[6,9] := -0.10753838;
      W_f[6,10] := 0.04849733;
      W_f[6,11] := -0.13716577;
      W_f[6,12] := 0.18706277;
      W_f[6,13] := -0.04876500;
      W_f[6,14] := 0.05665914;
      W_f[6,15] := -0.11948875;
      W_f[6,16] := -0.20568089;
      W_f[6,17] := -0.11067722;
      W_f[6,18] := -0.01706523;
      W_f[6,19] := -0.19956405;
      W_f[6,20] := -0.05881590;
      W_f[6,21] := 0.01174473;
      W_f[6,22] := -0.01817511;
      W_f[6,23] := 0.13952067;
      W_f[6,24] := 0.01716661;
      W_f[6,25] := 0.00872201;
      W_f[6,26] := 0.01365177;
      W_f[6,27] := 0.05093091;
      W_f[6,28] := -0.04843360;
      W_f[6,29] := -0.17431611;
      W_f[6,30] := -0.06636601;
      W_f[6,31] := -0.12669794;
      W_f[6,32] := 0.08169867;
      W_f[6,33] := 0.07502075;
      W_f[6,34] := 0.10079820;
      W_f[6,35] := 0.16185181;
      W_f[6,36] := -0.01285993;
      W_f[6,37] := -0.09518798;
      W_f[6,38] := -0.01886093;
      W_f[6,39] := -0.09482189;
      W_f[7,0] := 0.06969649;
      W_f[7,1] := 0.01038889;
      W_f[7,2] := 0.03716235;
      W_f[7,3] := 0.06842206;
      W_f[7,4] := 0.01828078;
      W_f[7,5] := 0.01142439;
      W_f[7,6] := -0.02572686;
      W_f[7,7] := -0.12288462;
      W_f[7,8] := -0.09727559;
      W_f[7,9] := 0.03457938;
      W_f[7,10] := 0.01338098;
      W_f[7,11] := -0.07754584;
      W_f[7,12] := 0.02478097;
      W_f[7,13] := -0.02415841;
      W_f[7,14] := -0.08689038;
      W_f[7,15] := -0.02232468;
      W_f[7,16] := 0.02237098;
      W_f[7,17] := -0.05418597;
      W_f[7,18] := 0.11298978;
      W_f[7,19] := 0.04869708;
      W_f[7,20] := -0.08651334;
      W_f[7,21] := 0.03297888;
      W_f[7,22] := -0.13389592;
      W_f[7,23] := 0.01270740;
      W_f[7,24] := -0.09401032;
      W_f[7,25] := 0.05024431;
      W_f[7,26] := -0.05931729;
      W_f[7,27] := 0.03168266;
      W_f[7,28] := 0.02225967;
      W_f[7,29] := 0.41531193;
      W_f[7,30] := -0.10573386;
      W_f[7,31] := -0.00634464;
      W_f[7,32] := 0.06730103;
      W_f[7,33] := -0.12398792;
      W_f[7,34] := 0.08676559;
      W_f[7,35] := 0.07915390;
      W_f[7,36] := -0.01929375;
      W_f[7,37] := 0.10289415;
      W_f[7,38] := -0.09580568;
      W_f[7,39] := 0.08953527;
      W_f[8,0] := 0.02770795;
      W_f[8,1] := 0.06031844;
      W_f[8,2] := -0.10150912;
      W_f[8,3] := 0.01504861;
      W_f[8,4] := -0.09168597;
      W_f[8,5] := 0.06771890;
      W_f[8,6] := -0.09644016;
      W_f[8,7] := 0.07058930;
      W_f[8,8] := 0.09084498;
      W_f[8,9] := 0.01001659;
      W_f[8,10] := -0.03256565;
      W_f[8,11] := -0.06310728;
      W_f[8,12] := -0.00573729;
      W_f[8,13] := 0.04646058;
      W_f[8,14] := -0.19100875;
      W_f[8,15] := -0.18868707;
      W_f[8,16] := 0.04595396;
      W_f[8,17] := -0.10153048;
      W_f[8,18] := -0.02347394;
      W_f[8,19] := 0.21639474;
      W_f[8,20] := -0.00608159;
      W_f[8,21] := -0.04918477;
      W_f[8,22] := 0.05360698;
      W_f[8,23] := -0.12926535;
      W_f[8,24] := 0.76762730;
      W_f[8,25] := 0.58518553;
      W_f[8,26] := -0.25098571;
      W_f[8,27] := 0.00410500;
      W_f[8,28] := 0.09514121;
      W_f[8,29] := -0.10038645;
      W_f[8,30] := 0.06295488;
      W_f[8,31] := -0.13594523;
      W_f[8,32] := 0.02679093;
      W_f[8,33] := -0.03734758;
      W_f[8,34] := 0.52519041;
      W_f[8,35] := 0.05038884;
      W_f[8,36] := -0.06236759;
      W_f[8,37] := 0.26230776;
      W_f[8,38] := -0.01351269;
      W_f[8,39] := 0.01838806;
      W_f[9,0] := 0.04727024;
      W_f[9,1] := 0.06008144;
      W_f[9,2] := -0.17861722;
      W_f[9,3] := -0.13905220;
      W_f[9,4] := 0.08026224;
      W_f[9,5] := -0.09055442;
      W_f[9,6] := 0.25250804;
      W_f[9,7] := 0.23927838;
      W_f[9,8] := -0.32988387;
      W_f[9,9] := -0.04884759;
      W_f[9,10] := -0.12125893;
      W_f[9,11] := -0.13363348;
      W_f[9,12] := 0.09538809;
      W_f[9,13] := 0.05378080;
      W_f[9,14] := 0.09597345;
      W_f[9,15] := 0.12151758;
      W_f[9,16] := 0.03207635;
      W_f[9,17] := 0.06979542;
      W_f[9,18] := 0.09580968;
      W_f[9,19] := 0.06583982;
      W_f[9,20] := 0.13815849;
      W_f[9,21] := -0.06946179;
      W_f[9,22] := 0.16799128;
      W_f[9,23] := -0.00493719;
      W_f[9,24] := -0.01021040;
      W_f[9,25] := 0.19830738;
      W_f[9,26] := -0.04321670;
      W_f[9,27] := 0.07314714;
      W_f[9,28] := -0.03591828;
      W_f[9,29] := 0.05154232;
      W_f[9,30] := -0.00456730;
      W_f[9,31] := 0.04409983;
      W_f[9,32] := -0.09231672;
      W_f[9,33] := 0.00690090;
      W_f[9,34] := 0.11396845;
      W_f[9,35] := 0.16058512;
      W_f[9,36] := -0.03188523;
      W_f[9,37] := -0.09661251;
      W_f[9,38] := 0.05787448;
      W_f[9,39] := 0.05807154;
      W_f[10,0] := 0.13345452;
      W_f[10,1] := 0.03274992;
      W_f[10,2] := -0.11242057;
      W_f[10,3] := -0.16067596;
      W_f[10,4] := 0.32250786;
      W_f[10,5] := -0.03652117;
      W_f[10,6] := -0.06048543;
      W_f[10,7] := 0.01128129;
      W_f[10,8] := -0.04134291;
      W_f[10,9] := 0.01602995;
      W_f[10,10] := 0.14861420;
      W_f[10,11] := -0.18624187;
      W_f[10,12] := 0.39872715;
      W_f[10,13] := 0.01673330;
      W_f[10,14] := -0.10627669;
      W_f[10,15] := 0.12056257;
      W_f[10,16] := 0.15113747;
      W_f[10,17] := -0.02927510;
      W_f[10,18] := -0.60066605;
      W_f[10,19] := -0.16866782;
      W_f[10,20] := -0.13441689;
      W_f[10,21] := 0.16711260;
      W_f[10,22] := 0.52250689;
      W_f[10,23] := -0.16760729;
      W_f[10,24] := -0.36896053;
      W_f[10,25] := -0.39812967;
      W_f[10,26] := 0.01471901;
      W_f[10,27] := -0.20327935;
      W_f[10,28] := -0.27292597;
      W_f[10,29] := 0.00824856;
      W_f[10,30] := 0.32700816;
      W_f[10,31] := -0.42109445;
      W_f[10,32] := -0.04604208;
      W_f[10,33] := 0.18438594;
      W_f[10,34] := 0.17093237;
      W_f[10,35] := -0.54145467;
      W_f[10,36] := -0.01911491;
      W_f[10,37] := -0.63746744;
      W_f[10,38] := 0.12846465;
      W_f[10,39] := -0.02683445;
      W_f[11,0] := -0.05971623;
      W_f[11,1] := 0.04910073;
      W_f[11,2] := 0.00890621;
      W_f[11,3] := 0.02669080;
      W_f[11,4] := -0.02135999;
      W_f[11,5] := 0.00178900;
      W_f[11,6] := 0.06730210;
      W_f[11,7] := -0.02445485;
      W_f[11,8] := 0.02154719;
      W_f[11,9] := 0.08513900;
      W_f[11,10] := -0.00957253;
      W_f[11,11] := 0.03944959;
      W_f[11,12] := 0.05303077;
      W_f[11,13] := 0.06797016;
      W_f[11,14] := 0.02574354;
      W_f[11,15] := 0.03408344;
      W_f[11,16] := -0.01919723;
      W_f[11,17] := -0.04070394;
      W_f[11,18] := 0.09808615;
      W_f[11,19] := 0.04076335;
      W_f[11,20] := 0.11645951;
      W_f[11,21] := 0.03692744;
      W_f[11,22] := -0.18985488;
      W_f[11,23] := -0.38257152;
      W_f[11,24] := -0.01752078;
      W_f[11,25] := 0.02452086;
      W_f[11,26] := 0.12240800;
      W_f[11,27] := 0.04160059;
      W_f[11,28] := -0.03000608;
      W_f[11,29] := -0.02825012;
      W_f[11,30] := 0.05161938;
      W_f[11,31] := 0.07235450;
      W_f[11,32] := -0.16787599;
      W_f[11,33] := 0.16893364;
      W_f[11,34] := 0.15554214;
      W_f[11,35] := -0.09419880;
      W_f[11,36] := -0.16331309;
      W_f[11,37] := -0.17827170;
      W_f[11,38] := 0.00083755;
      W_f[11,39] := 0.18259366;
      W_f[12,0] := -0.00770674;
      W_f[12,1] := 0.01958637;
      W_f[12,2] := -0.12229911;
      W_f[12,3] := 0.01299630;
      W_f[12,4] := -0.17465268;
      W_f[12,5] := 0.05698227;
      W_f[12,6] := -0.01131545;
      W_f[12,7] := -0.00422412;
      W_f[12,8] := -0.05034647;
      W_f[12,9] := 0.11572821;
      W_f[12,10] := -0.02485367;
      W_f[12,11] := -0.16879559;
      W_f[12,12] := -0.01365941;
      W_f[12,13] := -0.13796245;
      W_f[12,14] := 0.17325994;
      W_f[12,15] := -0.21148756;
      W_f[12,16] := 0.02845169;
      W_f[12,17] := 0.01354862;
      W_f[12,18] := -0.06274647;
      W_f[12,19] := -0.04003462;
      W_f[12,20] := 0.03278174;
      W_f[12,21] := 0.00519902;
      W_f[12,22] := -0.09380586;
      W_f[12,23] := 0.00667400;
      W_f[12,24] := 0.35337117;
      W_f[12,25] := 0.14751016;
      W_f[12,26] := 0.00971417;
      W_f[12,27] := 0.07586189;
      W_f[12,28] := 0.14462680;
      W_f[12,29] := -0.31107655;
      W_f[12,30] := 0.04906277;
      W_f[12,31] := -0.00521361;
      W_f[12,32] := -0.11651076;
      W_f[12,33] := 0.18232529;
      W_f[12,34] := 0.10977875;
      W_f[12,35] := -0.04999982;
      W_f[12,36] := -0.02277171;
      W_f[12,37] := -0.11629970;
      W_f[12,38] := -0.15014403;
      W_f[12,39] := -0.36427626;
      W_f[13,0] := -0.07062645;
      W_f[13,1] := -0.01207117;
      W_f[13,2] := -0.01288252;
      W_f[13,3] := 0.08112531;
      W_f[13,4] := -0.05332141;
      W_f[13,5] := 0.02898212;
      W_f[13,6] := -0.00224098;
      W_f[13,7] := 0.01993622;
      W_f[13,8] := 0.09566581;
      W_f[13,9] := -0.04889251;
      W_f[13,10] := -0.04912526;
      W_f[13,11] := -0.13804390;
      W_f[13,12] := -0.01942297;
      W_f[13,13] := 0.11708253;
      W_f[13,14] := 0.02629174;
      W_f[13,15] := -0.13945958;
      W_f[13,16] := -0.07286663;
      W_f[13,17] := -0.00936016;
      W_f[13,18] := -0.04328432;
      W_f[13,19] := -0.06046297;
      W_f[13,20] := -0.05109459;
      W_f[13,21] := 0.15283288;
      W_f[13,22] := -0.12800813;
      W_f[13,23] := -0.05418115;
      W_f[13,24] := 1.21206045;
      W_f[13,25] := 1.06606841;
      W_f[13,26] := -0.12827054;
      W_f[13,27] := -0.05296004;
      W_f[13,28] := 0.05082989;
      W_f[13,29] := 0.05279872;
      W_f[13,30] := -0.07762696;
      W_f[13,31] := -0.01807367;
      W_f[13,32] := 0.17315291;
      W_f[13,33] := 0.07421064;
      W_f[13,34] := 0.86849803;
      W_f[13,35] := 0.36573714;
      W_f[13,36] := -0.02259749;
      W_f[13,37] := 0.49192774;
      W_f[13,38] := -0.01003352;
      W_f[13,39] := 0.02914682;
      W_f[14,0] := -0.07975613;
      W_f[14,1] := 0.13247445;
      W_f[14,2] := -0.06722725;
      W_f[14,3] := 0.02443754;
      W_f[14,4] := 0.08127654;
      W_f[14,5] := 0.14814174;
      W_f[14,6] := 0.17534903;
      W_f[14,7] := 0.24142317;
      W_f[14,8] := -0.07938510;
      W_f[14,9] := 0.01944998;
      W_f[14,10] := -0.24030949;
      W_f[14,11] := 0.10943807;
      W_f[14,12] := 0.06249294;
      W_f[14,13] := -0.04712199;
      W_f[14,14] := 0.11892370;
      W_f[14,15] := 0.05002554;
      W_f[14,16] := 0.04903306;
      W_f[14,17] := 0.13278966;
      W_f[14,18] := -0.09704322;
      W_f[14,19] := -0.01522042;
      W_f[14,20] := 0.19409117;
      W_f[14,21] := 0.07847122;
      W_f[14,22] := 0.01956500;
      W_f[14,23] := -0.02513723;
      W_f[14,24] := -0.46761647;
      W_f[14,25] := -0.27084172;
      W_f[14,26] := 0.22476183;
      W_f[14,27] := 0.01039684;
      W_f[14,28] := 0.03313066;
      W_f[14,29] := 0.49718869;
      W_f[14,30] := 0.00785091;
      W_f[14,31] := 0.31502768;
      W_f[14,32] := 0.10209885;
      W_f[14,33] := 0.25726008;
      W_f[14,34] := 0.04868334;
      W_f[14,35] := -0.06811446;
      W_f[14,36] := -0.26499566;
      W_f[14,37] := -0.11457458;
      W_f[14,38] := -0.13219638;
      W_f[14,39] := -0.26006001;
      W_f[15,0] := -0.04342698;
      W_f[15,1] := 0.03330465;
      W_f[15,2] := -0.15716130;
      W_f[15,3] := 0.11637414;
      W_f[15,4] := 0.00085861;
      W_f[15,5] := 0.04937513;
      W_f[15,6] := -0.03373890;
      W_f[15,7] := 0.10901977;
      W_f[15,8] := -0.04058894;
      W_f[15,9] := -0.08138926;
      W_f[15,10] := -0.00654504;
      W_f[15,11] := 0.14907332;
      W_f[15,12] := -0.06752129;
      W_f[15,13] := -0.05585046;
      W_f[15,14] := 0.09911564;
      W_f[15,15] := -0.00484761;
      W_f[15,16] := 0.01454945;
      W_f[15,17] := -0.01109192;
      W_f[15,18] := -0.03362690;
      W_f[15,19] := 0.02557084;
      W_f[15,20] := -0.08767220;
      W_f[15,21] := 0.00880393;
      W_f[15,22] := -0.01261946;
      W_f[15,23] := -0.01694086;
      W_f[15,24] := 0.07210945;
      W_f[15,25] := 0.02202999;
      W_f[15,26] := -0.13439135;
      W_f[15,27] := -0.00877297;
      W_f[15,28] := 0.00261266;
      W_f[15,29] := -0.07274885;
      W_f[15,30] := -0.06177441;
      W_f[15,31] := 0.01014565;
      W_f[15,32] := -0.02689987;
      W_f[15,33] := -0.08880914;
      W_f[15,34] := -0.23302077;
      W_f[15,35] := -0.07694786;
      W_f[15,36] := -0.01976549;
      W_f[15,37] := -0.11379942;
      W_f[15,38] := 0.20449123;
      W_f[15,39] := -0.11346783;
      W_f[16,0] := -0.06895591;
      W_f[16,1] := -0.03991242;
      W_f[16,2] := 0.07949317;
      W_f[16,3] := -0.13159253;
      W_f[16,4] := 0.02148025;
      W_f[16,5] := -0.01628318;
      W_f[16,6] := 0.04405365;
      W_f[16,7] := 0.01672859;
      W_f[16,8] := -0.04237301;
      W_f[16,9] := 0.13518204;
      W_f[16,10] := -0.02853350;
      W_f[16,11] := -0.07497366;
      W_f[16,12] := -0.19952835;
      W_f[16,13] := -0.04520181;
      W_f[16,14] := 0.18698026;
      W_f[16,15] := -0.22438036;
      W_f[16,16] := -0.06152339;
      W_f[16,17] := -0.18698199;
      W_f[16,18] := 0.04692160;
      W_f[16,19] := 0.40312031;
      W_f[16,20] := 0.04334361;
      W_f[16,21] := -0.07279057;
      W_f[16,22] := 0.23739196;
      W_f[16,23] := 0.03972591;
      W_f[16,24] := -0.18138212;
      W_f[16,25] := -0.08058426;
      W_f[16,26] := -0.05819782;
      W_f[16,27] := -0.11114023;
      W_f[16,28] := -0.04217467;
      W_f[16,29] := -0.03431201;
      W_f[16,30] := -0.01802105;
      W_f[16,31] := 0.08157863;
      W_f[16,32] := -0.14787740;
      W_f[16,33] := 0.04127774;
      W_f[16,34] := -0.34828743;
      W_f[16,35] := -0.13249493;
      W_f[16,36] := 0.04573625;
      W_f[16,37] := -0.19219472;
      W_f[16,38] := -0.09764937;
      W_f[16,39] := -0.13595925;
      W_f[17,0] := 0.10454150;
      W_f[17,1] := -0.03026063;
      W_f[17,2] := -0.00496180;
      W_f[17,3] := -0.16523391;
      W_f[17,4] := 0.07944248;
      W_f[17,5] := 0.01923002;
      W_f[17,6] := 0.06903784;
      W_f[17,7] := 0.26167822;
      W_f[17,8] := -0.18167816;
      W_f[17,9] := 0.04501382;
      W_f[17,10] := -0.02101610;
      W_f[17,11] := -0.10886642;
      W_f[17,12] := 0.19678667;
      W_f[17,13] := -0.05605550;
      W_f[17,14] := -0.20257466;
      W_f[17,15] := -0.08576699;
      W_f[17,16] := -0.02321531;
      W_f[17,17] := 0.20090720;
      W_f[17,18] := 0.11825493;
      W_f[17,19] := 0.11430272;
      W_f[17,20] := 0.02607111;
      W_f[17,21] := 0.42574841;
      W_f[17,22] := 0.16701193;
      W_f[17,23] := -0.19879840;
      W_f[17,24] := -0.42272153;
      W_f[17,25] := -0.44768301;
      W_f[17,26] := 0.10922134;
      W_f[17,27] := -0.29530475;
      W_f[17,28] := -0.10366873;
      W_f[17,29] := 0.46814829;
      W_f[17,30] := 0.03179893;
      W_f[17,31] := 0.15740445;
      W_f[17,32] := 0.25256434;
      W_f[17,33] := 0.19541481;
      W_f[17,34] := 0.01293977;
      W_f[17,35] := -0.07509716;
      W_f[17,36] := -0.17786877;
      W_f[17,37] := 0.06767861;
      W_f[17,38] := -0.05990307;
      W_f[17,39] := 0.81737500;
      W_f[18,0] := 0.34308577;
      W_f[18,1] := -0.08164916;
      W_f[18,2] := -0.40619314;
      W_f[18,3] := -0.19120942;
      W_f[18,4] := 0.08112001;
      W_f[18,5] := 0.04640236;
      W_f[18,6] := -0.11047447;
      W_f[18,7] := 0.19122396;
      W_f[18,8] := -0.02393395;
      W_f[18,9] := 0.08837730;
      W_f[18,10] := -0.07884857;
      W_f[18,11] := 0.02850161;
      W_f[18,12] := -0.03546034;
      W_f[18,13] := 0.07510088;
      W_f[18,14] := -0.00984286;
      W_f[18,15] := -0.13105999;
      W_f[18,16] := 0.22273166;
      W_f[18,17] := -0.02799993;
      W_f[18,18] := 0.00293659;
      W_f[18,19] := 0.20137461;
      W_f[18,20] := -0.04015484;
      W_f[18,21] := 0.10801568;
      W_f[18,22] := -0.04284893;
      W_f[18,23] := 0.05038416;
      W_f[18,24] := -0.08880481;
      W_f[18,25] := -0.15249683;
      W_f[18,26] := 0.13808288;
      W_f[18,27] := 0.00168190;
      W_f[18,28] := -0.04924094;
      W_f[18,29] := -0.00257390;
      W_f[18,30] := -0.02845873;
      W_f[18,31] := 0.02481154;
      W_f[18,32] := -0.02671171;
      W_f[18,33] := 0.04705410;
      W_f[18,34] := -0.40709364;
      W_f[18,35] := 0.08703322;
      W_f[18,36] := -0.07230620;
      W_f[18,37] := 0.12350995;
      W_f[18,38] := 0.15746908;
      W_f[18,39] := -0.11168111;
      W_f[19,0] := 0.06964543;
      W_f[19,1] := 0.16963933;
      W_f[19,2] := -0.10727351;
      W_f[19,3] := -0.06463805;
      W_f[19,4] := -0.08993005;
      W_f[19,5] := -0.00428362;
      W_f[19,6] := 0.06947535;
      W_f[19,7] := 0.11149358;
      W_f[19,8] := -0.02489202;
      W_f[19,9] := -0.06382310;
      W_f[19,10] := 0.04778928;
      W_f[19,11] := -0.03058575;
      W_f[19,12] := -0.05471989;
      W_f[19,13] := 0.11426779;
      W_f[19,14] := -0.06128769;
      W_f[19,15] := -0.05338088;
      W_f[19,16] := 0.03729861;
      W_f[19,17] := -0.00755690;
      W_f[19,18] := 0.02605470;
      W_f[19,19] := -0.06562791;
      W_f[19,20] := -0.13053814;
      W_f[19,21] := 0.13839112;
      W_f[19,22] := 0.09563566;
      W_f[19,23] := -0.14636911;
      W_f[19,24] := 0.73496079;
      W_f[19,25] := 0.61294490;
      W_f[19,26] := -0.12774414;
      W_f[19,27] := -0.07314135;
      W_f[19,28] := 0.08495209;
      W_f[19,29] := 0.19162866;
      W_f[19,30] := -0.01792493;
      W_f[19,31] := -0.02980782;
      W_f[19,32] := -0.04641222;
      W_f[19,33] := 0.20514162;
      W_f[19,34] := 0.23501983;
      W_f[19,35] := 0.26531109;
      W_f[19,36] := 0.01960006;
      W_f[19,37] := 0.32003433;
      W_f[19,38] := -0.03473999;
      W_f[19,39] := 0.09161426;
      W_f[20,0] := -0.08032684;
      W_f[20,1] := 0.03764400;
      W_f[20,2] := 0.04910958;
      W_f[20,3] := -0.04065493;
      W_f[20,4] := -0.08581132;
      W_f[20,5] := 0.04799789;
      W_f[20,6] := -0.00371342;
      W_f[20,7] := -0.17297724;
      W_f[20,8] := 0.19704738;
      W_f[20,9] := 0.04339945;
      W_f[20,10] := -0.04020957;
      W_f[20,11] := -0.25716218;
      W_f[20,12] := -0.20699285;
      W_f[20,13] := 0.09457813;
      W_f[20,14] := 0.06039828;
      W_f[20,15] := -0.03535963;
      W_f[20,16] := 0.02864634;
      W_f[20,17] := -0.01065293;
      W_f[20,18] := -0.07240798;
      W_f[20,19] := -0.10301849;
      W_f[20,20] := 0.05020411;
      W_f[20,21] := 0.08534832;
      W_f[20,22] := 0.12433831;
      W_f[20,23] := -0.13624057;
      W_f[20,24] := 1.08051872;
      W_f[20,25] := 1.20131576;
      W_f[20,26] := -0.22155558;
      W_f[20,27] := 0.05610569;
      W_f[20,28] := 0.01186761;
      W_f[20,29] := -0.22767767;
      W_f[20,30] := 0.28332528;
      W_f[20,31] := 0.18194595;
      W_f[20,32] := 0.06990111;
      W_f[20,33] := -0.05628906;
      W_f[20,34] := 1.20703590;
      W_f[20,35] := 0.39179030;
      W_f[20,36] := 0.00589672;
      W_f[20,37] := 0.60747558;
      W_f[20,38] := 0.25271067;
      W_f[20,39] := 0.29734689;
      W_f[21,0] := 0.35368252;
      W_f[21,1] := -0.17104757;
      W_f[21,2] := -0.19149908;
      W_f[21,3] := -0.34622109;
      W_f[21,4] := 0.05045484;
      W_f[21,5] := -0.02223583;
      W_f[21,6] := 0.15965690;
      W_f[21,7] := 0.09061475;
      W_f[21,8] := -0.22678624;
      W_f[21,9] := 0.18206379;
      W_f[21,10] := 0.12876000;
      W_f[21,11] := 0.14537387;
      W_f[21,12] := 0.19264843;
      W_f[21,13] := -0.06770154;
      W_f[21,14] := 0.20032635;
      W_f[21,15] := -0.07122288;
      W_f[21,16] := -0.17053159;
      W_f[21,17] := 0.20213194;
      W_f[21,18] := -0.14164022;
      W_f[21,19] := 0.90530616;
      W_f[21,20] := -0.02790328;
      W_f[21,21] := -0.01270169;
      W_f[21,22] := -0.06040226;
      W_f[21,23] := 0.14147551;
      W_f[21,24] := -0.42720819;
      W_f[21,25] := -0.34853670;
      W_f[21,26] := 0.00898072;
      W_f[21,27] := -0.03843918;
      W_f[21,28] := -0.05057624;
      W_f[21,29] := 0.03018636;
      W_f[21,30] := -0.08073866;
      W_f[21,31] := 0.00180846;
      W_f[21,32] := -0.24050622;
      W_f[21,33] := -0.17357877;
      W_f[21,34] := 0.06599429;
      W_f[21,35] := -0.26927751;
      W_f[21,36] := -0.01186142;
      W_f[21,37] := -0.22601065;
      W_f[21,38] := 0.07210836;
      W_f[21,39] := 0.92559713;
      W_f[22,0] := 0.10358280;
      W_f[22,1] := 0.06531076;
      W_f[22,2] := -0.10848440;
      W_f[22,3] := -0.07142127;
      W_f[22,4] := 0.05051512;
      W_f[22,5] := 0.00920350;
      W_f[22,6] := -0.06956775;
      W_f[22,7] := 0.00521163;
      W_f[22,8] := -0.05201783;
      W_f[22,9] := 0.15847443;
      W_f[22,10] := -0.05266168;
      W_f[22,11] := -0.15218990;
      W_f[22,12] := -0.18027736;
      W_f[22,13] := 0.03990427;
      W_f[22,14] := 0.04980688;
      W_f[22,15] := 0.10445115;
      W_f[22,16] := -0.22353676;
      W_f[22,17] := 0.02329998;
      W_f[22,18] := -0.05035058;
      W_f[22,19] := -0.04183880;
      W_f[22,20] := -0.11790692;
      W_f[22,21] := 0.08537365;
      W_f[22,22] := 0.16631745;
      W_f[22,23] := -0.04788234;
      W_f[22,24] := 0.84037429;
      W_f[22,25] := 0.86304367;
      W_f[22,26] := -0.01927258;
      W_f[22,27] := 0.11064481;
      W_f[22,28] := 0.00307026;
      W_f[22,29] := -0.06691942;
      W_f[22,30] := 0.11506618;
      W_f[22,31] := -0.18648425;
      W_f[22,32] := 0.19806179;
      W_f[22,33] := -0.04705258;
      W_f[22,34] := 0.88099205;
      W_f[22,35] := 0.20989533;
      W_f[22,36] := 0.03750733;
      W_f[22,37] := 0.33899969;
      W_f[22,38] := 0.11258788;
      W_f[22,39] := 0.05194032;
      W_f[23,0] := 0.10712738;
      W_f[23,1] := 0.06521086;
      W_f[23,2] := -0.11553867;
      W_f[23,3] := 0.02760724;
      W_f[23,4] := 0.00875419;
      W_f[23,5] := 0.06495681;
      W_f[23,6] := -0.08853875;
      W_f[23,7] := 0.20240821;
      W_f[23,8] := -0.23240013;
      W_f[23,9] := -0.15616068;
      W_f[23,10] := 0.04585300;
      W_f[23,11] := 0.05213043;
      W_f[23,12] := 0.01046342;
      W_f[23,13] := -0.01021028;
      W_f[23,14] := -0.01159339;
      W_f[23,15] := -0.00385108;
      W_f[23,16] := -0.10526726;
      W_f[23,17] := -0.02686086;
      W_f[23,18] := 0.04239808;
      W_f[23,19] := 0.04591978;
      W_f[23,20] := 0.00747242;
      W_f[23,21] := 0.00471720;
      W_f[23,22] := 0.06718684;
      W_f[23,23] := 0.02261411;
      W_f[23,24] := -0.46556318;
      W_f[23,25] := -0.38187489;
      W_f[23,26] := -0.15911962;
      W_f[23,27] := -0.04183679;
      W_f[23,28] := 0.00261953;
      W_f[23,29] := 0.20375709;
      W_f[23,30] := 0.04742884;
      W_f[23,31] := -0.04061780;
      W_f[23,32] := -0.27790031;
      W_f[23,33] := -0.33751869;
      W_f[23,34] := -0.22227961;
      W_f[23,35] := -0.22620232;
      W_f[23,36] := 0.01848036;
      W_f[23,37] := 0.06976109;
      W_f[23,38] := 0.17023148;
      W_f[23,39] := 0.06424201;
      W_f[24,0] := -0.13167678;
      W_f[24,1] := 0.04912768;
      W_f[24,2] := 0.08014815;
      W_f[24,3] := -0.02571813;
      W_f[24,4] := -0.09035327;
      W_f[24,5] := -0.02664648;
      W_f[24,6] := -0.01713989;
      W_f[24,7] := -0.06988919;
      W_f[24,8] := 0.08913397;
      W_f[24,9] := 0.06661738;
      W_f[24,10] := -0.01555318;
      W_f[24,11] := -0.07162424;
      W_f[24,12] := -0.06340355;
      W_f[24,13] := -0.00172007;
      W_f[24,14] := 0.10926212;
      W_f[24,15] := -0.08084438;
      W_f[24,16] := -0.05963473;
      W_f[24,17] := -0.00672480;
      W_f[24,18] := 0.01630116;
      W_f[24,19] := -0.25053534;
      W_f[24,20] := -0.09545689;
      W_f[24,21] := 0.07690240;
      W_f[24,22] := 0.10612939;
      W_f[24,23] := -0.16514739;
      W_f[24,24] := 1.03784764;
      W_f[24,25] := 0.88065898;
      W_f[24,26] := -0.03682305;
      W_f[24,27] := -0.00828455;
      W_f[24,28] := 0.05003088;
      W_f[24,29] := -0.04010022;
      W_f[24,30] := 0.05692153;
      W_f[24,31] := 0.18359843;
      W_f[24,32] := 0.34326431;
      W_f[24,33] := 0.10616989;
      W_f[24,34] := 1.03922319;
      W_f[24,35] := 0.36108708;
      W_f[24,36] := -0.02607207;
      W_f[24,37] := 0.46878794;
      W_f[24,38] := 0.06349315;
      W_f[24,39] := -0.07822424;
      W_f[25,0] := 0.09424307;
      W_f[25,1] := -0.07596510;
      W_f[25,2] := -0.02230152;
      W_f[25,3] := -0.02251400;
      W_f[25,4] := -0.08674552;
      W_f[25,5] := -0.03909100;
      W_f[25,6] := 0.02012826;
      W_f[25,7] := -0.19810320;
      W_f[25,8] := -0.03501223;
      W_f[25,9] := 0.07801583;
      W_f[25,10] := 0.12167831;
      W_f[25,11] := 0.02942345;
      W_f[25,12] := -0.03074818;
      W_f[25,13] := 0.18136154;
      W_f[25,14] := -0.07766207;
      W_f[25,15] := -0.11802950;
      W_f[25,16] := 0.09643847;
      W_f[25,17] := -0.00825175;
      W_f[25,18] := -0.01346704;
      W_f[25,19] := 0.14435892;
      W_f[25,20] := -0.09294306;
      W_f[25,21] := 0.24677505;
      W_f[25,22] := -0.00171631;
      W_f[25,23] := -0.05241786;
      W_f[25,24] := -0.62711388;
      W_f[25,25] := -0.86187011;
      W_f[25,26] := -0.02512074;
      W_f[25,27] := -0.12612289;
      W_f[25,28] := 0.02822581;
      W_f[25,29] := 0.17376989;
      W_f[25,30] := 0.14752750;
      W_f[25,31] := -0.03002137;
      W_f[25,32] := 0.11643431;
      W_f[25,33] := 0.12692985;
      W_f[25,34] := 0.09470735;
      W_f[25,35] := -0.08044017;
      W_f[25,36] := -0.02479267;
      W_f[25,37] := -0.05792825;
      W_f[25,38] := -0.19763654;
      W_f[25,39] := 0.10607097;
      W_f[26,0] := -0.03801338;
      W_f[26,1] := 0.12077316;
      W_f[26,2] := -0.00214674;
      W_f[26,3] := 0.08969341;
      W_f[26,4] := -0.05175069;
      W_f[26,5] := 0.09671398;
      W_f[26,6] := 0.05628202;
      W_f[26,7] := 0.00741576;
      W_f[26,8] := 0.09492744;
      W_f[26,9] := 0.04450374;
      W_f[26,10] := -0.12498721;
      W_f[26,11] := -0.06016764;
      W_f[26,12] := -0.02876252;
      W_f[26,13] := 0.07218547;
      W_f[26,14] := -0.00462019;
      W_f[26,15] := -0.20534116;
      W_f[26,16] := -0.01119605;
      W_f[26,17] := -0.02882672;
      W_f[26,18] := 0.29306915;
      W_f[26,19] := -0.08930067;
      W_f[26,20] := 0.11014070;
      W_f[26,21] := 0.01036068;
      W_f[26,22] := -0.03047423;
      W_f[26,23] := -0.01341770;
      W_f[26,24] := 0.71706861;
      W_f[26,25] := 0.82642710;
      W_f[26,26] := -0.03907864;
      W_f[26,27] := 0.03413987;
      W_f[26,28] := 0.07479441;
      W_f[26,29] := 0.11823042;
      W_f[26,30] := -0.01580876;
      W_f[26,31] := 0.13751128;
      W_f[26,32] := 0.04258600;
      W_f[26,33] := -0.00015547;
      W_f[26,34] := 0.03845869;
      W_f[26,35] := 0.14624235;
      W_f[26,36] := 0.05640004;
      W_f[26,37] := 0.24197158;
      W_f[26,38] := 0.05926150;
      W_f[26,39] := 0.00147703;
      W_f[27,0] := -0.41983348;
      W_f[27,1] := 0.04596116;
      W_f[27,2] := 0.50369281;
      W_f[27,3] := -0.24023004;
      W_f[27,4] := -0.12844686;
      W_f[27,5] := 0.08288544;
      W_f[27,6] := -0.04881310;
      W_f[27,7] := 0.13240901;
      W_f[27,8] := -0.23897819;
      W_f[27,9] := 0.17269602;
      W_f[27,10] := -0.23331153;
      W_f[27,11] := 0.09929879;
      W_f[27,12] := -0.05380810;
      W_f[27,13] := -0.22379196;
      W_f[27,14] := -0.01404754;
      W_f[27,15] := -0.17665520;
      W_f[27,16] := -0.23467498;
      W_f[27,17] := -0.03324463;
      W_f[27,18] := -0.29978797;
      W_f[27,19] := 0.18120803;
      W_f[27,20] := -0.07370343;
      W_f[27,21] := 0.05440885;
      W_f[27,22] := 0.09849205;
      W_f[27,23] := -0.12451717;
      W_f[27,24] := -0.39236844;
      W_f[27,25] := -0.29468319;
      W_f[27,26] := 0.12390357;
      W_f[27,27] := -0.26659656;
      W_f[27,28] := 0.00462124;
      W_f[27,29] := -0.05021441;
      W_f[27,30] := 0.12468525;
      W_f[27,31] := -0.17938502;
      W_f[27,32] := 0.00435782;
      W_f[27,33] := 0.05119968;
      W_f[27,34] := -0.55093455;
      W_f[27,35] := -0.29848784;
      W_f[27,36] := 0.08519112;
      W_f[27,37] := -0.24839489;
      W_f[27,38] := 0.36261120;
      W_f[27,39] := -0.06641769;
      W_f[28,0] := -0.06259385;
      W_f[28,1] := -0.01964230;
      W_f[28,2] := -0.11223387;
      W_f[28,3] := 0.06842343;
      W_f[28,4] := 0.04186076;
      W_f[28,5] := 0.11873946;
      W_f[28,6] := 0.08319110;
      W_f[28,7] := 0.03873431;
      W_f[28,8] := -0.07993847;
      W_f[28,9] := -0.04896510;
      W_f[28,10] := -0.13774043;
      W_f[28,11] := -0.20616460;
      W_f[28,12] := 0.06616147;
      W_f[28,13] := -0.01874916;
      W_f[28,14] := 0.03724797;
      W_f[28,15] := 0.00960479;
      W_f[28,16] := -0.02171122;
      W_f[28,17] := -0.00924961;
      W_f[28,18] := -0.00415419;
      W_f[28,19] := -0.21919148;
      W_f[28,20] := -0.12006514;
      W_f[28,21] := 0.10141461;
      W_f[28,22] := 0.04794988;
      W_f[28,23] := 0.01126605;
      W_f[28,24] := -0.01665904;
      W_f[28,25] := -0.00120305;
      W_f[28,26] := 0.01582476;
      W_f[28,27] := 0.15678771;
      W_f[28,28] := -0.03058264;
      W_f[28,29] := 0.10287163;
      W_f[28,30] := 0.02894953;
      W_f[28,31] := -0.13468033;
      W_f[28,32] := -0.20077161;
      W_f[28,33] := 0.18928961;
      W_f[28,34] := 0.01422058;
      W_f[28,35] := 0.03234510;
      W_f[28,36] := -0.04311192;
      W_f[28,37] := -0.08474723;
      W_f[28,38] := 0.06878947;
      W_f[28,39] := 0.13092239;
      W_f[29,0] := -0.23808074;
      W_f[29,1] := -0.33427835;
      W_f[29,2] := -0.18062195;
      W_f[29,3] := -0.44995224;
      W_f[29,4] := -0.47261029;
      W_f[29,5] := 0.04930299;
      W_f[29,6] := -0.14416015;
      W_f[29,7] := -0.16943012;
      W_f[29,8] := 0.11852527;
      W_f[29,9] := 0.10351186;
      W_f[29,10] := 0.08463526;
      W_f[29,11] := 0.09515283;
      W_f[29,12] := 0.04440456;
      W_f[29,13] := -0.09559766;
      W_f[29,14] := -0.00851051;
      W_f[29,15] := -0.03550709;
      W_f[29,16] := -0.06376176;
      W_f[29,17] := -0.04328245;
      W_f[29,18] := 0.05228878;
      W_f[29,19] := -0.04287386;
      W_f[29,20] := 0.17943747;
      W_f[29,21] := 0.15752576;
      W_f[29,22] := 0.25777707;
      W_f[29,23] := -0.07851151;
      W_f[29,24] := -0.01634266;
      W_f[29,25] := -0.04672897;
      W_f[29,26] := 0.16563641;
      W_f[29,27] := -0.14571881;
      W_f[29,28] := 0.30397785;
      W_f[29,29] := 0.07079765;
      W_f[29,30] := 0.06753556;
      W_f[29,31] := -0.13499920;
      W_f[29,32] := -0.00998395;
      W_f[29,33] := 0.06980532;
      W_f[29,34] := -0.01776855;
      W_f[29,35] := -0.05868817;
      W_f[29,36] := -0.02662778;
      W_f[29,37] := 0.21032780;
      W_f[29,38] := -0.02339596;
      W_f[29,39] := -0.06946197;
      W_f[30,0] := -0.08261926;
      W_f[30,1] := -0.09091716;
      W_f[30,2] := 0.03065251;
      W_f[30,3] := 0.03797822;
      W_f[30,4] := -0.01897933;
      W_f[30,5] := 0.02048461;
      W_f[30,6] := -0.05789832;
      W_f[30,7] := -0.09650940;
      W_f[30,8] := 0.02682795;
      W_f[30,9] := -0.04769692;
      W_f[30,10] := 0.01357674;
      W_f[30,11] := -0.19160482;
      W_f[30,12] := 0.08094538;
      W_f[30,13] := -0.02382125;
      W_f[30,14] := -0.02338882;
      W_f[30,15] := 0.06300223;
      W_f[30,16] := 0.09212611;
      W_f[30,17] := -0.11708011;
      W_f[30,18] := 0.05085100;
      W_f[30,19] := 0.11342009;
      W_f[30,20] := -0.02413465;
      W_f[30,21] := -0.01437216;
      W_f[30,22] := 0.00564185;
      W_f[30,23] := -0.06922011;
      W_f[30,24] := -0.29297990;
      W_f[30,25] := -0.23998971;
      W_f[30,26] := 0.00216557;
      W_f[30,27] := 0.00281825;
      W_f[30,28] := -0.04129997;
      W_f[30,29] := 0.16728577;
      W_f[30,30] := 0.03681864;
      W_f[30,31] := 0.05884687;
      W_f[30,32] := -0.07153721;
      W_f[30,33] := 0.14938165;
      W_f[30,34] := -0.11850394;
      W_f[30,35] := -0.18422285;
      W_f[30,36] := 0.04826922;
      W_f[30,37] := -0.00851108;
      W_f[30,38] := 0.14509185;
      W_f[30,39] := -0.11933939;
      W_f[31,0] := 0.08570898;
      W_f[31,1] := 0.06335066;
      W_f[31,2] := -0.08633077;
      W_f[31,3] := 0.04141757;
      W_f[31,4] := -0.04193645;
      W_f[31,5] := 0.10255765;
      W_f[31,6] := 0.10652506;
      W_f[31,7] := -0.19849022;
      W_f[31,8] := -0.07185815;
      W_f[31,9] := 0.20198317;
      W_f[31,10] := 0.22491492;
      W_f[31,11] := -0.04794567;
      W_f[31,12] := -0.03101581;
      W_f[31,13] := 0.06656876;
      W_f[31,14] := -0.10685236;
      W_f[31,15] := -0.02540462;
      W_f[31,16] := 0.00684258;
      W_f[31,17] := -0.03772927;
      W_f[31,18] := 0.05183686;
      W_f[31,19] := 0.09021188;
      W_f[31,20] := -0.03484273;
      W_f[31,21] := 0.09286161;
      W_f[31,22] := 0.06733710;
      W_f[31,23] := -0.06343131;
      W_f[31,24] := 0.50989604;
      W_f[31,25] := 0.42543718;
      W_f[31,26] := -0.15198684;
      W_f[31,27] := 0.04894760;
      W_f[31,28] := 0.01305311;
      W_f[31,29] := 0.15279900;
      W_f[31,30] := 0.27127236;
      W_f[31,31] := 0.03008500;
      W_f[31,32] := 0.28474066;
      W_f[31,33] := 0.05558186;
      W_f[31,34] := 0.46742201;
      W_f[31,35] := 0.05888501;
      W_f[31,36] := -0.07833006;
      W_f[31,37] := 0.25103787;
      W_f[31,38] := 0.04388468;
      W_f[31,39] := 0.02715803;
      W_g[0,0] := -0.12131844;
      W_g[0,1] := 0.12085552;
      W_g[0,2] := 0.08980677;
      W_g[0,3] := 0.17669852;
      W_g[0,4] := -0.17395604;
      W_g[0,5] := 0.05983386;
      W_g[0,6] := -0.12038706;
      W_g[0,7] := 0.10408965;
      W_g[0,8] := 0.04987235;
      W_g[0,9] := 0.05143051;
      W_g[0,10] := -0.10646743;
      W_g[0,11] := -0.23724760;
      W_g[0,12] := 0.19022150;
      W_g[0,13] := 0.04472460;
      W_g[0,14] := -0.07482351;
      W_g[0,15] := -0.17896613;
      W_g[0,16] := 0.01789535;
      W_g[0,17] := -0.08042584;
      W_g[0,18] := 0.01418886;
      W_g[0,19] := 0.08560449;
      W_g[0,20] := 0.12055533;
      W_g[0,21] := -0.09562387;
      W_g[0,22] := 0.10016913;
      W_g[0,23] := -0.01397176;
      W_g[0,24] := 0.16734384;
      W_g[0,25] := 0.16720419;
      W_g[0,26] := 0.25958651;
      W_g[0,27] := 0.25067577;
      W_g[0,28] := 0.20941940;
      W_g[0,29] := -0.08324938;
      W_g[0,30] := 0.00226516;
      W_g[0,31] := -0.16828296;
      W_g[0,32] := -0.05718424;
      W_g[0,33] := -0.11489945;
      W_g[0,34] := 0.39200705;
      W_g[0,35] := -0.02924966;
      W_g[0,36] := -0.07215840;
      W_g[0,37] := -0.00060382;
      W_g[0,38] := 0.00190298;
      W_g[0,39] := -0.10329624;
      W_g[1,0] := 0.25078791;
      W_g[1,1] := -0.09808160;
      W_g[1,2] := -0.02631936;
      W_g[1,3] := -0.04027300;
      W_g[1,4] := 0.18441203;
      W_g[1,5] := 0.41963693;
      W_g[1,6] := 0.51547539;
      W_g[1,7] := 0.03554025;
      W_g[1,8] := -0.07983816;
      W_g[1,9] := 0.02190001;
      W_g[1,10] := -0.00606993;
      W_g[1,11] := 0.06645570;
      W_g[1,12] := 0.04269591;
      W_g[1,13] := 0.02085278;
      W_g[1,14] := 0.00638806;
      W_g[1,15] := 0.13739663;
      W_g[1,16] := 0.08046133;
      W_g[1,17] := -0.13583119;
      W_g[1,18] := -0.00408393;
      W_g[1,19] := 0.00235980;
      W_g[1,20] := 0.56796187;
      W_g[1,21] := -0.02013912;
      W_g[1,22] := -0.07913697;
      W_g[1,23] := -0.02018822;
      W_g[1,24] := -0.10366332;
      W_g[1,25] := 0.05380014;
      W_g[1,26] := -0.04720289;
      W_g[1,27] := -0.09928206;
      W_g[1,28] := -0.05330637;
      W_g[1,29] := 0.03338305;
      W_g[1,30] := 0.13593376;
      W_g[1,31] := 0.03519171;
      W_g[1,32] := 0.05909251;
      W_g[1,33] := 0.05970544;
      W_g[1,34] := 0.06835675;
      W_g[1,35] := -0.06630721;
      W_g[1,36] := 0.13448878;
      W_g[1,37] := 0.03730081;
      W_g[1,38] := 0.07570644;
      W_g[1,39] := -0.10574443;
      W_g[2,0] := -0.15925199;
      W_g[2,1] := 0.09215169;
      W_g[2,2] := 0.18303214;
      W_g[2,3] := -0.08564852;
      W_g[2,4] := 0.07656058;
      W_g[2,5] := -0.00410216;
      W_g[2,6] := 0.21223526;
      W_g[2,7] := -0.13624576;
      W_g[2,8] := -0.06400398;
      W_g[2,9] := -0.12832262;
      W_g[2,10] := 0.12734218;
      W_g[2,11] := 0.03441266;
      W_g[2,12] := -0.05592468;
      W_g[2,13] := 0.09095973;
      W_g[2,14] := -0.10887443;
      W_g[2,15] := -0.07970205;
      W_g[2,16] := 0.00062569;
      W_g[2,17] := -0.05494741;
      W_g[2,18] := 0.01040240;
      W_g[2,19] := 0.04842303;
      W_g[2,20] := -0.01907582;
      W_g[2,21] := 0.42660147;
      W_g[2,22] := -0.11769458;
      W_g[2,23] := -0.09431285;
      W_g[2,24] := -0.10584085;
      W_g[2,25] := -0.25145948;
      W_g[2,26] := -0.03071128;
      W_g[2,27] := 0.22361481;
      W_g[2,28] := 0.05417244;
      W_g[2,29] := -0.05925388;
      W_g[2,30] := -0.08127954;
      W_g[2,31] := 0.06508211;
      W_g[2,32] := -0.00114283;
      W_g[2,33] := -0.08544528;
      W_g[2,34] := -0.21091597;
      W_g[2,35] := 0.13263747;
      W_g[2,36] := -0.21554339;
      W_g[2,37] := 0.10003000;
      W_g[2,38] := 0.01394136;
      W_g[2,39] := -0.00390853;
      W_g[3,0] := 0.20485403;
      W_g[3,1] := -0.11455492;
      W_g[3,2] := 0.18512601;
      W_g[3,3] := 0.18688123;
      W_g[3,4] := -0.21285971;
      W_g[3,5] := 0.07757265;
      W_g[3,6] := -0.20667188;
      W_g[3,7] := 0.06186296;
      W_g[3,8] := -0.30767784;
      W_g[3,9] := -0.13624844;
      W_g[3,10] := -0.17604175;
      W_g[3,11] := -0.01812170;
      W_g[3,12] := 0.59569001;
      W_g[3,13] := 0.08554336;
      W_g[3,14] := 0.30720758;
      W_g[3,15] := -0.47165588;
      W_g[3,16] := -0.31375375;
      W_g[3,17] := -0.31498158;
      W_g[3,18] := 0.05816992;
      W_g[3,19] := -0.03276125;
      W_g[3,20] := 0.11148553;
      W_g[3,21] := -0.45352960;
      W_g[3,22] := -0.43782380;
      W_g[3,23] := -0.11082695;
      W_g[3,24] := -0.20848672;
      W_g[3,25] := -0.12392744;
      W_g[3,26] := 0.04257244;
      W_g[3,27] := 0.16871507;
      W_g[3,28] := 0.11623926;
      W_g[3,29] := 0.06922457;
      W_g[3,30] := -0.45511082;
      W_g[3,31] := 1.14466596;
      W_g[3,32] := 0.04183885;
      W_g[3,33] := 0.45074558;
      W_g[3,34] := 0.02823192;
      W_g[3,35] := 0.01668284;
      W_g[3,36] := -0.08451141;
      W_g[3,37] := 0.19031323;
      W_g[3,38] := -0.11998753;
      W_g[3,39] := 0.70253503;
      W_g[4,0] := -0.08821924;
      W_g[4,1] := 0.22643130;
      W_g[4,2] := 0.21002994;
      W_g[4,3] := -0.20082740;
      W_g[4,4] := -0.00453639;
      W_g[4,5] := -0.08484363;
      W_g[4,6] := -0.06815410;
      W_g[4,7] := -0.02295598;
      W_g[4,8] := -0.18677296;
      W_g[4,9] := 0.01185095;
      W_g[4,10] := 0.41826287;
      W_g[4,11] := 0.05190533;
      W_g[4,12] := -0.15545513;
      W_g[4,13] := -0.14982492;
      W_g[4,14] := 0.01574554;
      W_g[4,15] := 0.18053719;
      W_g[4,16] := 0.03002386;
      W_g[4,17] := 0.02935749;
      W_g[4,18] := 0.02353674;
      W_g[4,19] := -0.02946706;
      W_g[4,20] := 0.04099213;
      W_g[4,21] := -0.11064263;
      W_g[4,22] := 0.06823131;
      W_g[4,23] := 0.29373077;
      W_g[4,24] := -0.01898101;
      W_g[4,25] := -0.02048161;
      W_g[4,26] := -0.26626879;
      W_g[4,27] := 0.26876929;
      W_g[4,28] := -0.01425563;
      W_g[4,29] := 0.22355153;
      W_g[4,30] := 0.26949978;
      W_g[4,31] := 0.26295567;
      W_g[4,32] := 0.16207495;
      W_g[4,33] := 0.00838947;
      W_g[4,34] := 0.21043131;
      W_g[4,35] := 0.00681238;
      W_g[4,36] := 0.01988858;
      W_g[4,37] := 0.13659397;
      W_g[4,38] := 0.11311906;
      W_g[4,39] := -0.04562292;
      W_g[5,0] := 0.17928106;
      W_g[5,1] := 0.26329628;
      W_g[5,2] := -0.10853200;
      W_g[5,3] := -0.09602788;
      W_g[5,4] := -0.16062686;
      W_g[5,5] := -0.06875742;
      W_g[5,6] := 0.14379244;
      W_g[5,7] := 0.05838383;
      W_g[5,8] := -0.13917951;
      W_g[5,9] := 0.05606813;
      W_g[5,10] := 0.02034150;
      W_g[5,11] := -0.01945914;
      W_g[5,12] := -0.18592170;
      W_g[5,13] := -0.11316089;
      W_g[5,14] := -0.16464360;
      W_g[5,15] := 0.02854693;
      W_g[5,16] := 0.00971764;
      W_g[5,17] := -0.06508735;
      W_g[5,18] := 0.00310314;
      W_g[5,19] := -0.14046571;
      W_g[5,20] := -0.23027138;
      W_g[5,21] := -0.20236713;
      W_g[5,22] := 0.02430346;
      W_g[5,23] := -0.14275949;
      W_g[5,24] := -0.09406747;
      W_g[5,25] := 0.21386193;
      W_g[5,26] := -0.03222166;
      W_g[5,27] := 0.01500143;
      W_g[5,28] := 0.11013638;
      W_g[5,29] := -0.07420376;
      W_g[5,30] := 0.00631831;
      W_g[5,31] := -0.13111025;
      W_g[5,32] := 0.00536069;
      W_g[5,33] := -0.05818216;
      W_g[5,34] := -0.17104428;
      W_g[5,35] := -0.05052703;
      W_g[5,36] := 0.15376194;
      W_g[5,37] := 0.09446555;
      W_g[5,38] := -0.02123900;
      W_g[5,39] := 0.10707947;
      W_g[6,0] := -0.18866111;
      W_g[6,1] := 0.12487285;
      W_g[6,2] := 0.02589516;
      W_g[6,3] := -0.09877703;
      W_g[6,4] := -0.08392680;
      W_g[6,5] := -0.03048542;
      W_g[6,6] := 0.07423776;
      W_g[6,7] := 0.09883864;
      W_g[6,8] := 0.08149955;
      W_g[6,9] := 0.15533857;
      W_g[6,10] := -0.10272066;
      W_g[6,11] := 0.18736395;
      W_g[6,12] := -0.24082580;
      W_g[6,13] := 0.01097316;
      W_g[6,14] := -0.01382545;
      W_g[6,15] := 0.03999422;
      W_g[6,16] := 0.14499241;
      W_g[6,17] := 0.10716019;
      W_g[6,18] := 0.01429422;
      W_g[6,19] := 0.21958458;
      W_g[6,20] := 0.34892666;
      W_g[6,21] := 0.16072913;
      W_g[6,22] := -0.03282092;
      W_g[6,23] := -0.00633068;
      W_g[6,24] := -0.39161780;
      W_g[6,25] := -0.20158361;
      W_g[6,26] := -0.03133341;
      W_g[6,27] := -0.09530033;
      W_g[6,28] := 0.16384017;
      W_g[6,29] := 0.05612209;
      W_g[6,30] := 0.04608196;
      W_g[6,31] := 0.17323117;
      W_g[6,32] := -0.09182145;
      W_g[6,33] := -0.13467614;
      W_g[6,34] := -0.33367291;
      W_g[6,35] := -0.06024042;
      W_g[6,36] := 0.04037794;
      W_g[6,37] := -0.14040722;
      W_g[6,38] := -0.00377652;
      W_g[6,39] := 0.22859706;
      W_g[7,0] := 0.30623785;
      W_g[7,1] := 0.22891158;
      W_g[7,2] := 0.05204437;
      W_g[7,3] := 0.09328783;
      W_g[7,4] := 0.08432135;
      W_g[7,5] := -0.03246771;
      W_g[7,6] := 0.06265932;
      W_g[7,7] := -0.10986651;
      W_g[7,8] := 0.27611876;
      W_g[7,9] := -0.04993419;
      W_g[7,10] := -0.05604714;
      W_g[7,11] := -0.04595119;
      W_g[7,12] := -0.05060242;
      W_g[7,13] := -0.01598648;
      W_g[7,14] := 0.17354257;
      W_g[7,15] := 0.11727922;
      W_g[7,16] := -0.01031275;
      W_g[7,17] := 0.08838559;
      W_g[7,18] := -0.18819259;
      W_g[7,19] := 0.08691938;
      W_g[7,20] := 0.02175990;
      W_g[7,21] := -0.01114948;
      W_g[7,22] := -0.01792710;
      W_g[7,23] := 0.01326630;
      W_g[7,24] := 0.03426804;
      W_g[7,25] := 0.23651482;
      W_g[7,26] := 0.00880161;
      W_g[7,27] := 0.07044864;
      W_g[7,28] := -0.11657553;
      W_g[7,29] := -0.10108893;
      W_g[7,30] := -0.00445770;
      W_g[7,31] := 0.06863080;
      W_g[7,32] := -0.00541675;
      W_g[7,33] := -0.02590487;
      W_g[7,34] := 0.04817338;
      W_g[7,35] := 0.05935349;
      W_g[7,36] := -0.02825072;
      W_g[7,37] := 0.02169201;
      W_g[7,38] := 0.04781851;
      W_g[7,39] := -0.00979924;
      W_g[8,0] := -0.00056170;
      W_g[8,1] := 0.09928103;
      W_g[8,2] := -0.03647884;
      W_g[8,3] := -0.11951732;
      W_g[8,4] := -0.00163588;
      W_g[8,5] := -0.02342502;
      W_g[8,6] := 0.02331413;
      W_g[8,7] := 0.10044318;
      W_g[8,8] := -0.02542515;
      W_g[8,9] := 0.16847059;
      W_g[8,10] := 0.03315528;
      W_g[8,11] := 0.01159255;
      W_g[8,12] := 0.02168436;
      W_g[8,13] := 0.07067128;
      W_g[8,14] := 0.25364098;
      W_g[8,15] := -0.15877020;
      W_g[8,16] := 0.11872134;
      W_g[8,17] := -0.05331764;
      W_g[8,18] := -0.03777300;
      W_g[8,19] := 0.17292042;
      W_g[8,20] := 0.06789102;
      W_g[8,21] := -0.05720007;
      W_g[8,22] := 0.13237606;
      W_g[8,23] := -0.28390497;
      W_g[8,24] := 0.02519086;
      W_g[8,25] := -0.01009906;
      W_g[8,26] := -0.31023392;
      W_g[8,27] := 0.02227520;
      W_g[8,28] := 0.08983584;
      W_g[8,29] := 0.01240572;
      W_g[8,30] := 0.12657896;
      W_g[8,31] := -0.28511786;
      W_g[8,32] := 0.03818220;
      W_g[8,33] := 0.03446925;
      W_g[8,34] := -0.08904101;
      W_g[8,35] := -0.02425133;
      W_g[8,36] := -0.12229283;
      W_g[8,37] := -0.04048497;
      W_g[8,38] := -0.16955297;
      W_g[8,39] := 0.01971084;
      W_g[9,0] := 0.19825646;
      W_g[9,1] := 0.15505151;
      W_g[9,2] := 0.18824823;
      W_g[9,3] := 0.05656092;
      W_g[9,4] := -0.11205027;
      W_g[9,5] := 0.01548184;
      W_g[9,6] := -0.26724932;
      W_g[9,7] := 0.06024139;
      W_g[9,8] := 0.19550920;
      W_g[9,9] := 0.09395395;
      W_g[9,10] := -0.00923733;
      W_g[9,11] := 0.28975904;
      W_g[9,12] := -0.11834054;
      W_g[9,13] := 0.01023313;
      W_g[9,14] := -0.09161735;
      W_g[9,15] := -0.09301599;
      W_g[9,16] := 0.01594188;
      W_g[9,17] := -0.07896575;
      W_g[9,18] := -0.07530534;
      W_g[9,19] := -0.06356308;
      W_g[9,20] := -0.14556308;
      W_g[9,21] := 0.35489818;
      W_g[9,22] := -0.10316110;
      W_g[9,23] := -0.03947277;
      W_g[9,24] := 0.06387684;
      W_g[9,25] := -0.05773838;
      W_g[9,26] := -0.13109356;
      W_g[9,27] := -0.40293059;
      W_g[9,28] := 0.20684175;
      W_g[9,29] := 0.34316665;
      W_g[9,30] := 0.04913993;
      W_g[9,31] := 0.13192397;
      W_g[9,32] := 0.11378421;
      W_g[9,33] := 0.13727243;
      W_g[9,34] := -0.16840093;
      W_g[9,35] := 0.23456278;
      W_g[9,36] := 0.07689143;
      W_g[9,37] := 0.02866838;
      W_g[9,38] := -0.04906642;
      W_g[9,39] := 0.00189616;
      W_g[10,0] := 0.09864533;
      W_g[10,1] := 0.02665105;
      W_g[10,2] := -0.07577279;
      W_g[10,3] := 0.31387433;
      W_g[10,4] := 0.10285930;
      W_g[10,5] := 0.00906804;
      W_g[10,6] := 0.08912777;
      W_g[10,7] := -0.14490779;
      W_g[10,8] := 0.01400164;
      W_g[10,9] := -0.30717424;
      W_g[10,10] := 0.07055619;
      W_g[10,11] := -0.62748581;
      W_g[10,12] := 0.21564768;
      W_g[10,13] := -0.07443854;
      W_g[10,14] := -0.24998751;
      W_g[10,15] := 0.00295377;
      W_g[10,16] := -0.03179332;
      W_g[10,17] := 0.21825644;
      W_g[10,18] := -0.00976076;
      W_g[10,19] := -0.11549558;
      W_g[10,20] := 0.00315555;
      W_g[10,21] := 0.19182777;
      W_g[10,22] := 0.17524354;
      W_g[10,23] := -0.07308983;
      W_g[10,24] := -0.12984170;
      W_g[10,25] := 0.07283737;
      W_g[10,26] := 0.07790703;
      W_g[10,27] := -0.10306653;
      W_g[10,28] := -0.06413930;
      W_g[10,29] := 0.14150777;
      W_g[10,30] := 0.08703817;
      W_g[10,31] := -0.19606562;
      W_g[10,32] := -0.03046606;
      W_g[10,33] := 0.11359414;
      W_g[10,34] := 0.09200487;
      W_g[10,35] := -0.29436204;
      W_g[10,36] := 0.01480583;
      W_g[10,37] := -0.14805350;
      W_g[10,38] := 0.37741283;
      W_g[10,39] := 0.33747074;
      W_g[11,0] := 0.30691084;
      W_g[11,1] := 0.22507285;
      W_g[11,2] := -0.05586467;
      W_g[11,3] := -0.02278013;
      W_g[11,4] := -0.16402608;
      W_g[11,5] := -0.12950912;
      W_g[11,6] := 0.02949622;
      W_g[11,7] := 0.17381540;
      W_g[11,8] := -0.25788903;
      W_g[11,9] := 0.07214717;
      W_g[11,10] := 0.23979028;
      W_g[11,11] := 0.06327691;
      W_g[11,12] := -0.06549240;
      W_g[11,13] := 0.27871069;
      W_g[11,14] := 0.01952578;
      W_g[11,15] := 0.01537968;
      W_g[11,16] := -0.00508708;
      W_g[11,17] := 0.08779414;
      W_g[11,18] := -0.03233203;
      W_g[11,19] := -0.06247540;
      W_g[11,20] := 0.12738970;
      W_g[11,21] := -0.20136435;
      W_g[11,22] := -0.12966998;
      W_g[11,23] := -0.56388378;
      W_g[11,24] := -0.14447659;
      W_g[11,25] := -0.18179278;
      W_g[11,26] := 0.17201598;
      W_g[11,27] := 0.10523865;
      W_g[11,28] := 0.08958710;
      W_g[11,29] := -0.05589786;
      W_g[11,30] := -0.09582882;
      W_g[11,31] := 0.27669013;
      W_g[11,32] := -0.04552330;
      W_g[11,33] := 0.01918150;
      W_g[11,34] := 0.06293701;
      W_g[11,35] := -0.22501966;
      W_g[11,36] := -0.06364831;
      W_g[11,37] := -0.20046265;
      W_g[11,38] := 0.02329997;
      W_g[11,39] := -0.23204710;
      W_g[12,0] := 0.06894288;
      W_g[12,1] := 0.02977384;
      W_g[12,2] := -0.27906618;
      W_g[12,3] := 0.17588335;
      W_g[12,4] := 0.03122274;
      W_g[12,5] := -0.00869676;
      W_g[12,6] := 0.02498548;
      W_g[12,7] := 0.15665044;
      W_g[12,8] := -0.23465285;
      W_g[12,9] := -0.02305496;
      W_g[12,10] := 0.03085731;
      W_g[12,11] := -0.06395327;
      W_g[12,12] := 0.21618837;
      W_g[12,13] := -0.17170039;
      W_g[12,14] := 0.06037929;
      W_g[12,15] := 0.11929530;
      W_g[12,16] := -0.01636845;
      W_g[12,17] := -0.09329034;
      W_g[12,18] := -0.49559087;
      W_g[12,19] := 0.05422232;
      W_g[12,20] := -0.01635499;
      W_g[12,21] := 0.10374246;
      W_g[12,22] := -0.08315807;
      W_g[12,23] := 0.10288428;
      W_g[12,24] := 0.10813106;
      W_g[12,25] := 0.09857040;
      W_g[12,26] := 0.04437799;
      W_g[12,27] := -0.06397744;
      W_g[12,28] := -0.03081079;
      W_g[12,29] := 0.07190378;
      W_g[12,30] := -0.12962900;
      W_g[12,31] := 0.03743947;
      W_g[12,32] := -0.09458277;
      W_g[12,33] := -0.06948329;
      W_g[12,34] := -0.32606724;
      W_g[12,35] := -0.13728699;
      W_g[12,36] := 0.01340251;
      W_g[12,37] := 0.08566734;
      W_g[12,38] := -0.05628554;
      W_g[12,39] := -0.31428364;
      W_g[13,0] := -0.04341206;
      W_g[13,1] := 0.01232883;
      W_g[13,2] := 0.01258724;
      W_g[13,3] := 0.11650011;
      W_g[13,4] := -0.05845366;
      W_g[13,5] := -0.02547886;
      W_g[13,6] := -0.14294159;
      W_g[13,7] := -0.00287156;
      W_g[13,8] := 0.04528259;
      W_g[13,9] := -0.03991419;
      W_g[13,10] := -0.04396502;
      W_g[13,11] := -0.13575317;
      W_g[13,12] := 0.19402504;
      W_g[13,13] := -0.01273516;
      W_g[13,14] := 0.00092753;
      W_g[13,15] := -0.08336857;
      W_g[13,16] := -0.02212642;
      W_g[13,17] := -0.03646492;
      W_g[13,18] := -0.01780297;
      W_g[13,19] := -0.02802462;
      W_g[13,20] := 0.16785975;
      W_g[13,21] := 0.09308389;
      W_g[13,22] := -0.05633133;
      W_g[13,23] := 0.01729810;
      W_g[13,24] := -0.12873031;
      W_g[13,25] := -0.06776203;
      W_g[13,26] := -0.01449728;
      W_g[13,27] := 0.45830390;
      W_g[13,28] := -0.25314638;
      W_g[13,29] := -0.08932091;
      W_g[13,30] := -0.10103022;
      W_g[13,31] := -0.14912573;
      W_g[13,32] := -0.03426053;
      W_g[13,33] := 0.03538388;
      W_g[13,34] := -0.12175231;
      W_g[13,35] := -0.11719010;
